(* IEC 61131-3 sources: PLC-IsaVODE/PLC-IsaVODE/samples/plc-programs, 701 files *)

(* ---- 250-building.IEC ---- *)
(*@PROPERTIES_EX@
TYPE: DATA_TYPE
LOCALE: 0
*)
(* ------------------------------------------- *)

TYPE oscat_TIMER_EVENT_DATA :
  STRUCT
	TYP          : BYTE;
	CHANNEL      : BYTE;
	DAY          : BYTE;
	START        : UDINT;
	DURATION     : TIME;
	LAND         : BYTE;
	LOR          : BYTE;
	LAST         : UDINT;
  END_STRUCT;
END_TYPE

TYPE
  oscat_TIMER_EVENT           : ARRAY [0..63]    OF oscat_TIMER_EVENT_DATA;
END_TYPE

(* ------------------------------------------- *)

TYPE
  oscat_T_AVG24         	  : ARRAY [0..47]   OF INT;

  oscat_TP4_qn                : ARRAY [0..3]    OF BOOL;

  oscat_bsa_X                 : ARRAY [0..2]    OF BYTE;
  oscat_blind_scene_array     : ARRAY [0..15]   OF oscat_bsa_X;

END_TYPE

(* ---- 731-WORLD_WEATHER.ST ---- *)
TYPE
  oscat_STRING30              : STRING;
  oscat_STRING250             : STRING;
  oscat_STRING8               : STRING;
  oscat_STRING60               : STRING;
  oscat_STRING3               : STRING;
  oscat_STRING10               : STRING;
END_TYPE

TYPE
  oscat_IP_FIFO128_DATA  : ARRAY [1..128] OF BYTE;
  oscat_Mailbox  : ARRAY [1..16] OF BYTE;

  oscat_IP_FIFO_DATA :
  STRUCT
	X       : oscat_IP_FIFO128_DATA; (* IP_ID FIFO Speicher          *)
	Y       : oscat_IP_FIFO128_DATA; (* IP_ID Z�hler                 *)
	ID      : BYTE;                  (* h�chste vergabene id         *)
	MAX_ID  : BYTE;                  (* maximal Anmeldungen pro ID   *)
    INIT    : BOOL;                  (* Initialisierung durchgef�hrt *)
	EMPTY   : BOOL;                  (* FIFO leer                    *)
	FULL    : BOOL;                  (* FIFO voll                    *)
	TOP     : INT;                   (* maximale anzahl in FIFO      *)
	NW      : INT;                   (* Schreibzeiger                *)
	NR      : INT;                   (* Lesezeiger                   *)
  END_STRUCT;

  oscat_IP_C:
  STRUCT
  	C_MODE:			BYTE;          		(*W Mode: TCP/UCP AKTIV/PASSIV                               *)
	C_PORT:         WORD;          		(*W Portnummer                                               *)
	C_IP:           DWORD;         		(*W IP-Adresse gepackt wwxxyyzz = www.xxx.yyy.zzz            *)
    C_STATE:        BYTE;          		(*R Verbindungsstatus ON/OFF + Flanke ON/OFF                 *)
	C_ENABLE:       BOOL;          		(*W Freigabe f�r Connect                                     *)
    R_OBSERVE:      BOOL;          		(*W Empfang ueberwachen                                      *)
    TIME_RESET:     BOOL;          		(*W Alle Timer ruecksetzen                                   *)
	ERROR:          DWORD;         		(*R vvwwxxyy (vv = CON_ERROR, ww = SEN_ERROR, xx = REC_ERROR *)
    FIFO:           oscat_IP_FIFO_DATA; (*I IP FIFO Struktur                                         *)
	MAILBOX:		oscat_Mailbox;		(*I Mailbox: Datenbereich f�r Bausteindatenaustausch         *)
  END_STRUCT;

  oscat_XML_CONTROL:
  STRUCT
    COMMAND:             WORD;            (*W                 *)
    WATCHDOG:            TIME;            (*W                 *)
    START_POS:           UINT;            (*W                 *)
    STOP_POS:            UINT;            (*W                 *)
    COUNT:               UINT;            (*R                 *)
    TYP:                 INT;             (*R                 *)
    LEVEL:               UINT;            (*R                 *)
    PATH:                oscat_STRING250; (*R                 *)
    ELEMENT:             oscat_STRING250; (*R                 *)
    ATTRIBUTE:           oscat_STRING250; (*R                 *)
    VALUE:               oscat_STRING250; (*R                 *)
    BLOCK1_START:        UINT;            (*R                 *)
    BLOCK1_STOP:         UINT;            (*R                 *)
    BLOCK2_START:        UINT;            (*R                 *)
    BLOCK2_STOP:         UINT;            (*R                 *)
  END_STRUCT;

  (* --------- WORLD WEATHER --------- *)

  oscat_WORLD_WEATHER_CUR :
  STRUCT
	OBSERVATION_TIME : oscat_STRING8;
	TEMP_C           : INT;
	WEATHER_CODE     : INT;
	WEATHER_DESC 	 : oscat_STRING60;
	WEATHER_ICON     : INT;
	WIND_SPEED_MILES : INT;
	WIND_SPEED_KMPH  : INT;
	WIND_DIR_DEGREE  : INT;
	WIND_DIR16POINT  : oscat_STRING3;
	PRECIPMM         : REAL;
	HUMIDITY         : INT;
	VISIBILITY       : INT;
	PRESSURE         : INT;
	CLOUDOVER        : INT;
  END_STRUCT;

  oscat_WORLD_WEATHER_DAY :
  STRUCT
	DATE_OF_DAY      : oscat_STRING10;
	TEMP_MAX_C       : INT;
	TEMP_MAX_F       : INT;
	TEMP_MIN_C       : INT;
	TEMP_MIN_F       : INT;
	WIND_SPEED_MILES : INT;
	WIND_SPEED_KMPH  : INT;
	WIND_DIR_DEGREE  : INT;
	WIND_DIR16POINT  : oscat_STRING3;
	WEATHER_CODE     : INT;
	WEATHER_DESC     : oscat_STRING60;
	WEATHER_ICON     : INT;
	PRECIPMM         : REAL;
  END_STRUCT;

  oscat_WORLD_WEATHER_DAY_ARR : ARRAY [0..4] OF oscat_WORLD_WEATHER_DAY;

  oscat_WORLD_WEATHER_DATA :
  STRUCT
	CUR : oscat_WORLD_WEATHER_CUR;
	DAY : oscat_WORLD_WEATHER_DAY_ARR;
  END_STRUCT;

  oscat_WORLD_WEATHER_aI0_41 : ARRAY[0..41] OF INT;

END_TYPE

TYPE
  oscat_NW_BUF_LONG  : ARRAY [0..4095] OF BYTE;

  oscat_NETWORK_BUFFER :
  STRUCT
    SIZE   : UINT;
    BUFFER : oscat_NW_BUF_LONG;
  END_STRUCT;

END_TYPE

FUNCTION_BLOCK WORLD_WEATHER_Block

	VAR_INPUT
		ACTIVATE :	BOOL;
		LATITUDE :	REAL;
		LONGITUDE :	REAL;
		KEY :	oscat_STRING30;
	END_VAR

	VAR_OUTPUT
		BUSY :	BOOL;
		DONE :	BOOL;
		ERROR_C :	DWORD;
		ERROR_T :	BYTE;
	END_VAR

	VAR_IN_OUT
		IP_C :	oscat_IP_C;
		S_BUF :	oscat_NETWORK_BUFFER;
		R_BUF :	oscat_NETWORK_BUFFER;
		WW :	oscat_WORLD_WEATHER_DATA;
	END_VAR

	VAR
		CHK_REAL :	CHK_REAL;
		REAL_TO_STRF :	REAL_TO_STRF;
		URL_DATA :	oscat_url;
		DNS_CLIENT :	DNS_CLIENT;
		HTTP_GET :	HTTP_GET;
		CPB :	CSV_PARSER_BUF;
		STRING_TO_URL :	STRING_TO_URL;
		FLOAT_TO_REAL :	FLOAT_TO_REAL;
		last_state :	BOOL;
		value_int :	INT;
		value_real :	REAL;
		v_real :	REAL;
		state :	INT;
		url_str :	oscat_STRING250;
		offset :	UDINT;
		size :	INT;
		sep :	BYTE;
		cnt :	INT;
		day :	INT;
		idx :	INT;
		run :	BYTE;
		result :	BYTE;
		value :	oscat_STRING250;
		DEC_TO_INT :	DEC_TO_INT;
		pos :	INT;
	END_VAR

	CASE state OF

	00:
		IF ACTIVATE AND NOT last_state THEN
			state := 20;
			DONE := FALSE;
			BUSY := TRUE;
			ERROR_C := DWORD#0;
			ERROR_T := BYTE#0;
		END_IF;

	20:
		REAL_TO_STRF(IN:=LATITUDE,N:=6,D:='.');
		url_str := CONCAT('http://free.worldweatheronline.com/feed/weather.ashx?q=',REAL_TO_STRF.REAL_TO_STRF);
		url_str := CONCAT(url_str,',');
		REAL_TO_STRF(IN:=LONGITUDE,N:=6,D:='.');
		url_str := CONCAT(url_str,REAL_TO_STRF.REAL_TO_STRF);
		url_str := CONCAT(url_str,'&format=csv&num_of_days=5&key=');
		url_str := CONCAT(url_str,key);

		STRING_TO_URL(STR:=url_str, DEFAULT_PROTOCOL:='', DEFAULT_PATH:='' );
		URL_DATA:=STRING_TO_URL.STRING_TO_URL;

		state := 40;

	40:
		IF DNS_CLIENT.DONE THEN
			state := 60;
		ELSIF (DNS_CLIENT.ERROR > DWORD#00) THEN
			ERROR_C := DNS_CLIENT.ERROR;
			ERROR_T := BYTE#01;
			state   := 100;
		END_IF;

	60:
		IF HTTP_GET.DONE THEN
			sep := BYTE#0;
			idx := 0;
			day := 0;
			cnt := 0;
			OFFSET := UINT_TO_UDINT(HTTP_GET.BODY_START);
			size := UINT_TO_INT(HTTP_GET.BODY_STOP);
			run := BYTE#1;
			state := 80;

		ELSIF (HTTP_GET.ERROR > DWORD#00) THEN
			ERROR_C := HTTP_GET.ERROR;
			ERROR_T := BYTE#02;
			state := 100;
		END_IF;

	80:	IF run = BYTE#0 THEN
			run := BYTE#1;
			IF result = BYTE#1 OR result = BYTE#2 THEN
				value_int := 0;
				value_real := 0.0;
				IF LEN(value) <= 20 THEN
					FLOAT_TO_REAL(FLT:=value);
					v_real := FLOAT_TO_REAL.FLOAT_TO_REAL;
					CHK_REAL(X := v_real);
					IF CHK_REAL.CHK_REAL = BYTE#0 THEN
						value_real := v_real;
						value_int := REAL_TO_INT(value_real);
					END_IF;
				END_IF;
				cnt := cnt + 1;
				IF cnt >=8 AND cnt <= 87 THEN
					IF cnt > 22 THEN
						CASE idx OF
						00:	WW.DAY[day].DATE_OF_DAY := value;
						01:	WW.DAY[day].TEMP_MAX_C := value_int;
						02:	WW.DAY[day].TEMP_MAX_F := value_int;
						03:	WW.DAY[day].TEMP_MIN_C := value_int;
						04:	WW.DAY[day].TEMP_MIN_F := value_int;
						05:	WW.DAY[day].WIND_SPEED_MILES := value_int;
						06:	WW.DAY[day].WIND_SPEED_KMPH := value_int;
						07:	WW.DAY[day].WIND_DIR_DEGREE := value_int;
						08:	WW.DAY[day].WIND_DIR16POINT := value;
						09:	WW.DAY[day].WEATHER_CODE := value_int;
						10:	pos := FIND(value, '/wsymbol_');
							IF pos > 0 AND LEN(value) > pos + 13 THEN
								DEC_TO_INT(DEC:=MID(value,4,pos + 9));
								WW.DAY[day].WEATHER_ICON := DEC_TO_INT.DEC_TO_INT;
							ELSE
								WW.DAY[day].WEATHER_ICON := 0;
							END_IF;
						11:	WW.DAY[day].WEATHER_DESC := value;
						12:	WW.DAY[day].PRECIPMM := value_real;
						END_CASE;
						idx := idx + 1;
						IF idx > 12 THEN
							idx := 0;
							day := day + 1;
						END_IF;
					ELSE
						CASE cnt OF
						08:	sep := BYTE#44;
						09:	WW.CUR.OBSERVATION_TIME := value;
						10:	WW.CUR.TEMP_C := value_int;
						11:	WW.CUR.WEATHER_CODE := value_int;
						12:	pos := FIND(value, '/wsymbol_');
							IF pos > 0 AND LEN(value) > pos + 13 THEN
								DEC_TO_INT(DEC:=MID(value,4,pos + 9));
								WW.CUR.WEATHER_ICON := DEC_TO_INT.DEC_TO_INT;
							ELSE
								WW.CUR.WEATHER_ICON := 0;
							END_IF;
						13:	WW.CUR.WEATHER_DESC := value;
						14:	WW.CUR.WIND_SPEED_MILES := value_int;
						15:	WW.CUR.WIND_SPEED_KMPH := value_int;
						16:	WW.CUR.WIND_DIR_DEGREE := value_int;
						17:	WW.CUR.WIND_DIR16POINT := value;
						18:	WW.CUR.PRECIPMM := value_real;
						19:	WW.CUR.HUMIDITY := value_int;
						20:	WW.CUR.VISIBILITY := value_int;
						21:	WW.CUR.PRESSURE := value_int;
						22:	WW.CUR.CLOUDOVER := value_int;
						END_CASE;
					END_IF;
				END_IF;
			ELSIF result = BYTE#10 THEN
				DONE  := TRUE;
				run := BYTE#0;
				state := 100;
			END_IF;
		END_IF;

	100:
		IF (NOT HTTP_GET.DONE) THEN
			state := 0;
			BUSY := FALSE;
			DONE := ERROR_T = BYTE#0;
		END_IF;

	END_CASE;

	DNS_CLIENT.IP_C     := IP_C;
	DNS_CLIENT.S_BUF    := S_BUF;
	DNS_CLIENT.R_BUF    := R_BUF;
	DNS_CLIENT.DOMAIN   := URL_DATA.DOMAIN;
	DNS_CLIENT.IP4_DNS  := DWORD#00;
	DNS_CLIENT.ACTIVATE := state=40;
	DNS_CLIENT();
	IP_C  := DNS_CLIENT.IP_C;
	S_BUF := DNS_CLIENT.S_BUF;
	R_BUF := DNS_CLIENT.R_BUF;

	HTTP_GET.IP_C        := IP_C;
	HTTP_GET.S_BUF       := S_BUF;
	HTTP_GET.R_BUF       := R_BUF;
	HTTP_GET.IP4         := DNS_CLIENT.IP4;
	HTTP_GET.GET         := state=60;
	HTTP_GET.MODE        := BYTE#2;
	HTTP_GET.UNLOCK_BUF  := state=100;
	HTTP_GET.URL_DATA    := URL_DATA;
	HTTP_GET();
	IP_C     := HTTP_GET.IP_C;
	S_BUF    := HTTP_GET.S_BUF;
	R_BUF    := HTTP_GET.R_BUF;
	URL_DATA := HTTP_GET.URL_DATA;

	CPB(SEP:=sep,RUN:=run,OFFSET:=offset,VALUE:=value,PT:=R_BUF);
	run:=CPB.RUN;
	offset:=CPB.OFFSET;
	value:=CPB.VALUE;
	R_BUF:=CPB.PT;
	result:=CPB.RESULT;

	last_state := ACTIVATE;

END_FUNCTION_BLOCK

PROGRAM program0
	VAR
		ACTIVATE :	BOOL;
		LATITUDE :	REAL;
		LONGITUDE :	REAL;
		KEY :	oscat_STRING30;
		IP_C :	oscat_IP_C;
		S_BUF :	oscat_NETWORK_BUFFER;
		R_BUF :	oscat_NETWORK_BUFFER;
		WW :	oscat_WORLD_WEATHER_DATA;
		BUSY :	BOOL;
		DONE :	BOOL;
		ERROR_C :	DWORD;
		ERROR_T :	BYTE;

		func_block : WORLD_WEATHER_Block;
	END_VAR
	func_block.ACTIVATE := ACTIVATE;
	func_block.LATITUDE := LATITUDE;
	func_block.LONGITUDE := LONGITUDE;
	func_block.KEY := KEY;
	func_block.IP_C := IP_C;
	func_block.S_BUF := S_BUF;
	func_block.R_BUF := R_BUF;
	func_block.WW := WW;

	func_block();
	IP_C  := func_block.IP_C;
	S_BUF  := func_block.S_BUF;
	R_BUF  := func_block.R_BUF;
	WW  := func_block.WW;
	BUSY  := func_block.BUSY;
	DONE  := func_block.DONE;
	ERROR_C  := func_block.ERROR_C;
	ERROR_T  := func_block.ERROR_T;
END_PROGRAM

CONFIGURATION Config0
	RESOURCE Res0 ON PLC
		TASK task0(INTERVAL := T#20ms,PRIORITY := 0);
		PROGRAM instance0 WITH task0 : program0;
	END_RESOURCE
END_CONFIGURATION

(* ---- 733-YAHOO_WEATHER_ICON_OSCAT.ST ---- *)
TYPE
  oscat_STRING1               : STRING;
  oscat_STRING2               : STRING;
  oscat_STRING3               : STRING;
  oscat_STRING4               : STRING;
  oscat_STRING5               : STRING;
  oscat_STRING8               : STRING;
  oscat_STRING10              : STRING;
  oscat_STRING12            : STRING;
  oscat_STRING15            : STRING;
  oscat_STRING20            : STRING;
  oscat_STRING27            : STRING;
  oscat_STRING30            : STRING;
  oscat_STRING32            : STRING;
  oscat_STRING40            : STRING;
  oscat_STRING48            : STRING;
  oscat_STRING50            : STRING;
  oscat_STRING60            : STRING;
  oscat_STRING64            : STRING;
  oscat_STRING80            : STRING;
  oscat_STRING120            : STRING;
  oscat_STRING140            : STRING;
  oscat_STRING160            : STRING;
  oscat_STRING180            : STRING;
  oscat_STRING190            : STRING;
  oscat_STRING250            : STRING;
END_TYPE

TYPE
  oscat_IP_FIFO128_DATA  : ARRAY [1..128] OF BYTE;
  oscat_Mailbox  : ARRAY [1..16] OF BYTE;

  oscat_IP_FIFO_DATA :
  STRUCT
	X       : oscat_IP_FIFO128_DATA; (* IP_ID FIFO Speicher          *)
	Y       : oscat_IP_FIFO128_DATA; (* IP_ID Z�hler                 *)
	ID      : BYTE;                  (* h�chste vergabene id         *)
	MAX_ID  : BYTE;                  (* maximal Anmeldungen pro ID   *)
    INIT    : BOOL;                  (* Initialisierung durchgef�hrt *)
	EMPTY   : BOOL;                  (* FIFO leer                    *)
	FULL    : BOOL;                  (* FIFO voll                    *)
	TOP     : INT;                   (* maximale anzahl in FIFO      *)
	NW      : INT;                   (* Schreibzeiger                *)
	NR      : INT;                   (* Lesezeiger                   *)
  END_STRUCT;

  oscat_IP_C:
  STRUCT
  	C_MODE:			BYTE;          		(*W Mode: TCP/UCP AKTIV/PASSIV                               *)
	C_PORT:         WORD;          		(*W Portnummer                                               *)
	C_IP:           DWORD;         		(*W IP-Adresse gepackt wwxxyyzz = www.xxx.yyy.zzz            *)
    C_STATE:        BYTE;          		(*R Verbindungsstatus ON/OFF + Flanke ON/OFF                 *)
	C_ENABLE:       BOOL;          		(*W Freigabe f�r Connect                                     *)
    R_OBSERVE:      BOOL;          		(*W Empfang ueberwachen                                      *)
    TIME_RESET:     BOOL;          		(*W Alle Timer ruecksetzen                                   *)
	ERROR:          DWORD;         		(*R vvwwxxyy (vv = CON_ERROR, ww = SEN_ERROR, xx = REC_ERROR *)
    FIFO:           oscat_IP_FIFO_DATA; (*I IP FIFO Struktur                                         *)
	MAILBOX:		oscat_Mailbox;		(*I Mailbox: Datenbereich f�r Bausteindatenaustausch         *)
  END_STRUCT;

  oscat_XML_CONTROL:
  STRUCT
    COMMAND:             WORD;            (*W                 *)
    WATCHDOG:            TIME;            (*W                 *)
    START_POS:           UINT;            (*W                 *)
    STOP_POS:            UINT;            (*W                 *)
    COUNT:               UINT;            (*R                 *)
    TYP:                 INT;             (*R                 *)
    LEVEL:               UINT;            (*R                 *)
    PATH:                oscat_STRING250; (*R                 *)
    ELEMENT:             oscat_STRING250; (*R                 *)
    ATTRIBUTE:           oscat_STRING250; (*R                 *)
    VALUE:               oscat_STRING250; (*R                 *)
    BLOCK1_START:        UINT;            (*R                 *)
    BLOCK1_STOP:         UINT;            (*R                 *)
    BLOCK2_START:        UINT;            (*R                 *)
    BLOCK2_STOP:         UINT;            (*R                 *)
  END_STRUCT;

  (* --------- WORLD WEATHER --------- *)

  oscat_WORLD_WEATHER_CUR :
  STRUCT
	OBSERVATION_TIME : oscat_STRING8;
	TEMP_C           : INT;
	WEATHER_CODE     : INT;
	WEATHER_DESC 	 : oscat_STRING60;
	WEATHER_ICON     : INT;
	WIND_SPEED_MILES : INT;
	WIND_SPEED_KMPH  : INT;
	WIND_DIR_DEGREE  : INT;
	WIND_DIR16POINT  : oscat_STRING3;
	PRECIPMM         : REAL;
	HUMIDITY         : INT;
	VISIBILITY       : INT;
	PRESSURE         : INT;
	CLOUDOVER        : INT;
  END_STRUCT;

  oscat_WORLD_WEATHER_DAY :
  STRUCT
	DATE_OF_DAY      : oscat_STRING10;
	TEMP_MAX_C       : INT;
	TEMP_MAX_F       : INT;
	TEMP_MIN_C       : INT;
	TEMP_MIN_F       : INT;
	WIND_SPEED_MILES : INT;
	WIND_SPEED_KMPH  : INT;
	WIND_DIR_DEGREE  : INT;
	WIND_DIR16POINT  : oscat_STRING3;
	WEATHER_CODE     : INT;
	WEATHER_DESC     : oscat_STRING60;
	WEATHER_ICON     : INT;
	PRECIPMM         : REAL;
  END_STRUCT;

  oscat_WORLD_WEATHER_DAY_ARR : ARRAY [0..4] OF oscat_WORLD_WEATHER_DAY;

  oscat_WORLD_WEATHER_DATA :
  STRUCT
	CUR : oscat_WORLD_WEATHER_CUR;
	DAY : oscat_WORLD_WEATHER_DAY_ARR;
  END_STRUCT;

  oscat_WORLD_WEATHER_aI0_41 : ARRAY[0..41] OF INT;

  (* --------- WEATHER CHANNEL --------- *)
  oscat_YAHOO_WEATHER_DATA:
  STRUCT
    TIMETOLIVE:                 INT;              (* TIME TO LIVE: HOW LONG IN MINUTES THIS FEED SHOULD BE CACHED         *)
    LOCATION_CITY:              OSCAT_STRING40;   (* THE LOCATION OF THIS FORECAST: CITY: CITY NAME  *)
    LOCATION_REGION:            OSCAT_STRING20;   (* THE LOCATION OF THIS FORECAST: REGION: STATE, TERRITORY, OR REGION, IF GIVEN *)
    LOCATION_COUNTRY:           OSCAT_STRING20;    (* THE LOCATION OF THIS FORECAST: COUNTRY: TWO-CHARACTER COUNTRY CODE *)
    UNIT_TEMPERATURE:           OSCAT_STRING1;    (* TEMPERATURE: DEGREE UNITS, F FOR FAHRENHEIT OR C FOR CELSIUS *)
    UNIT_DISTANCE:              OSCAT_STRING2;    (* DISTANCE: UNITS FOR DISTANCE, MI FOR MILES OR KM FOR KILOMETERS *)
    UNIT_PRESSURE:              OSCAT_STRING2;    (* PRESSURE: UNITS OF BAROMETRIC PRESSURE, IN FOR POUNDS PER SQUARE INCH OR MB FOR MILLIBARS *)
    UNIT_SPEED:                 OSCAT_STRING4;    (* SPEED: UNITS OF SPEED, MPH FOR MILES PER HOUR OR KPH FOR KILOMETERS PER HOUR *)
    WIND_CHILL:                 INT;              (* FORECAST INFORMATION ABOUT WIND CHILL IN DEGREES *)
    WIND_DIRECTION:             INT;              (* FORECAST INFORMATION ABOUT WIND DIRECTION, IN DEGREES *)
    WIND_SPEED:                 REAL;             (* FORECAST INFORMATION ABOUT WIND SPEED, IN THE UNITS (MPH OR KPH)*)
    ATMOSPHERE_HUMIDITY:        INT;              (* FORECAST INFORMATION ABOUT CURRENT ATMOSPHERIC HUMIDITY: HUMIDITY, IN PERCENT  *)
    ATMOSPHERE_PRESSURE:        INT;              (* FORECAST INFORMATION ABOUT CURRENT ATMOSPHERIC PRESSURE: BAROMETRIC PRESSURE, IN THE UNITS (IN OR MB) *)
	ATMOSPHERE_VISIBILITY:      REAL;             (* FORECAST INFORMATION ABOUT CURRENT ATMOSPHERIC VISIBILITY, IN THE UNITS (MI OR KM) *)
	ATMOSPHERE_RISING:          INT;              (* FORECAST INFORMATION ABOUT RISING: STATE OF THE BAROMETRIC PRESSURE: STEADY (0), RISING (1), OR FALLING (2). (INTEGER: 0, 1, 2) *)
    ASTRONOMY_SUNRISE:          OSCAT_STRING10;   (* SUNRISE: TODAY'S SUNRISE TIME. THE TIME IS A STRING IN A LOCAL TIME FORMAT OF "H:MM AM/PM" *)
    ASTRONOMY_SUNSET:           OSCAT_STRING10;   (* SUNSET: TODAY'S SUNSET TIME. THE TIME IS A STRING IN A LOCAL TIME FORMAT OF "H:MM AM/PM", *)
    GEO_LATITUDE:               REAL;             (* THE LATITUDE OF THE LOCATION *)
    GEO_LONGITUDE:              REAL;             (* THE LONGITUDE OF THE LOCATION *)
    CUR_CONDITIONS_TEMP:        INT;              (* THE CURRENT WEATHER CONDITIONS: TEMP: THE CURRENT TEMPERATURE, IN THE UNITS (F OR C) *)
    CUR_CONDITIONS_TEXT:        OSCAT_STRING40;   (* THE CURRENT WEATHER CONDITIONS: TEXT: A TEXTUAL DESCRIPTION OF CONDITIONS *)
    CUR_CONDITIONS_CODE:        INT;              (* THE CURRENT WEATHER CONDITIONS: CODE: THE CONDITION CODE FOR THIS FORECAST *)
	CUR_CONDITIONS_ICON:        INT;			  (* THE CURRENT WEATHER CONDITIONS: ICON: THE CONDITION ICON FOR THIS FORECAST *)
    FORCAST_TODAY_LOW_TEMP:     INT;              (* THE FORCAST TODAY WEATHER CONDITIONS: THE FORECASTED LOW TEMPERATURE FOR THIS DAY IN THE UNITS (F OR C) *)
    FORCAST_TODAY_HIGH_TEMP:    INT;              (* THE FORCAST TODAY WEATHER CONDITIONS: THE FORECASTED HIGH TEMPERATURE FOR THIS DAY IN THE UNITS (F OR C) *)
    FORCAST_TODAY_TEXT:         OSCAT_STRING40;   (* THE FORCAST TODAY WEATHER CONDITIONS: TEXT: A TEXTUAL DESCRIPTION OF CONDITIONS *)
    FORCAST_TODAY_CODE:         INT;              (* THE CURRENT WEATHER CONDITIONS: CODE: THE CONDITION CODE FOR THIS FORECAST *)
	FORCAST_TODAY_ICON:         INT;			  (* THE CURRENT WEATHER CONDITIONS: ICON: THE CONDITION ICON FOR THIS FORECAST *)
    FORCAST_TOMORROW_LOW_TEMP:  INT;              (* THE FORCAST TOMORROW WEATHER CONDITIONS: THE FORECASTED LOW TEMPERATURE FOR THIS DAY IN THE UNITS (F OR C) *)
    FORCAST_TOMORROW_HIGH_TEMP: INT;              (* THE FORCAST TOMORROW WEATHER CONDITIONS: THE FORECASTED HIGH TEMPERATURE FOR THIS DAY IN THE UNITS (F OR C) *)
    FORCAST_TOMORROW_TEXT:      OSCAT_STRING40;   (* THE FORCAST TOMORROW WEATHER CONDITIONS: TEXT: A TEXTUAL DESCRIPTION OF CONDITIONS *)
    FORCAST_TOMORROW_CODE:      INT;              (* THE CURRENT WEATHER CONDITIONS: CODE: THE CONDITION CODE FOR THIS FORECAST *)
	FORCAST_TOMORROW_ICON:      INT;			  (* THE CURRENT WEATHER CONDITIONS: ICON: THE CONDITION ICON FOR THIS FORECAST *)
  END_STRUCT;

  oscat_YAHOO_WEATHER_aI0_48 : ARRAY[0..48] OF INT;

  oscat_IP2GEO_DATA:
  STRUCT
	STATE :				BOOL;			  (* STATE *)
	IP4 :				DWORD;			  (* IP-Adresse *)
    COUNTRY_CODE :		oscat_STRING2;    (*   *)
    COUNTRY_NAME :		oscat_STRING20;   (*   *)
    REGION_CODE :		oscat_STRING2;    (*   *)
    REGION_NAME :		oscat_STRING20;   (*   *)
    CITY :				oscat_STRING20;   (*   *)
    GEO_LATITUDE :		REAL;             (*   *)
    GEO_LONGITUDE :		REAL;             (*   *)
	TIME_ZONE_NAME :	oscat_STRING20;
	GMT_OFFSET :		INT;
	IS_DST :			BOOL;
  END_STRUCT;
END_TYPE

FUNCTION_BLOCK YAHOO_WEATHER_ICON_OSCAT_Block

	VAR_INPUT
		ACTIVATE :	BOOL;
	END_VAR

	VAR_IN_OUT
		YW :	oscat_YAHOO_WEATHER_DATA;
	END_VAR

	VAR
		act_last :	BOOL;
		x :	INT;
		init :	BOOL;
		dat :	oscat_YAHOO_WEATHER_aI0_48;
	END_VAR

	IF not init THEN
		init := TRUE;

		dat[00] := 4;
		dat[01] := 2;
		dat[02] := 2;
		dat[03] := 4;
		dat[04] := 17;
		dat[05] := 1;
		dat[06] := 3;
		dat[07] := 1;
		dat[08] := 2;
		dat[09] := 2;
		dat[10] := 2;
		dat[11] := 2;
		dat[12] := 2;
		dat[13] := 3;
		dat[14] := 3;
		dat[15] := 3;
		dat[16] := 3;
		dat[17] := 5;
		dat[18] := 3;
		dat[19] := 6;
		dat[20] := 7;
		dat[21] := 14;
		dat[22] := 8;
		dat[23] := 9;
		dat[24] := 9;
		dat[25] := 10;
		dat[26] := 9;
		dat[27] := 11;
		dat[28] := 12;
		dat[29] := 11;
		dat[30] := 12;
		dat[31] := 13;
		dat[32] := 14;
		dat[33] := 15;
		dat[34] := 16;
		dat[35] := 4;
		dat[36] := 14;
		dat[37] := 4;
		dat[38] := 17;
		dat[39] := 2;
		dat[40] := 2;
		dat[41] := 3;
		dat[42] := 3;
		dat[43] := 3;
		dat[44] := 12;
		dat[45] := 2;
		dat[46] := 3;
		dat[47] := 4;
		dat[48] := 0;
	END_IF;

	IF ACTIVATE AND act_last = FALSE THEN
		x := MIN(YW.CUR_CONDITIONS_CODE,48);
		YW.CUR_CONDITIONS_ICON := dat[x];
		x := MIN(YW.FORCAST_TODAY_CODE,48);
		YW.FORCAST_TODAY_ICON := dat[x];
		x := MIN(YW.FORCAST_TOMORROW_CODE,48);
		YW.FORCAST_TOMORROW_ICON := dat[x];
	END_IF;
	act_last := ACTIVATE;

END_FUNCTION_BLOCK

PROGRAM program0
	VAR
		ACTIVATE :	BOOL;
		YW :	oscat_YAHOO_WEATHER_DATA;

		func_block : YAHOO_WEATHER_ICON_OSCAT_Block;
	END_VAR
	func_block.ACTIVATE := ACTIVATE;
	func_block.YW := YW;

	func_block();
	YW  := func_block.YW;
END_PROGRAM

CONFIGURATION Config0
	RESOURCE Res0 ON PLC
		TASK task0(INTERVAL := T#20ms,PRIORITY := 0);
		PROGRAM instance0 WITH task0 : program0;
	END_RESOURCE
END_CONFIGURATION

(* ---- 737-YAHOO_WEATHER_DESC_GE.ST ---- *)
TYPE
  oscat_STRING1               : STRING;
  oscat_STRING2               : STRING;
  oscat_STRING3               : STRING;
  oscat_STRING4               : STRING;
  oscat_STRING5               : STRING;
  oscat_STRING8               : STRING;
  oscat_STRING10              : STRING;
  oscat_STRING12            : STRING;
  oscat_STRING15            : STRING;
  oscat_STRING20            : STRING;
  oscat_STRING27            : STRING;
  oscat_STRING30            : STRING;
  oscat_STRING32            : STRING;
  oscat_STRING40            : STRING;
  oscat_STRING48            : STRING;
  oscat_STRING50            : STRING;
  oscat_STRING60            : STRING;
  oscat_STRING64            : STRING;
  oscat_STRING80            : STRING;
  oscat_STRING120            : STRING;
  oscat_STRING140            : STRING;
  oscat_STRING160            : STRING;
  oscat_STRING180            : STRING;
  oscat_STRING190            : STRING;
  oscat_STRING250            : STRING;
END_TYPE

TYPE
  oscat_IP_FIFO128_DATA  : ARRAY [1..128] OF BYTE;
  oscat_Mailbox  : ARRAY [1..16] OF BYTE;

  oscat_IP_FIFO_DATA :
  STRUCT
	X       : oscat_IP_FIFO128_DATA; (* IP_ID FIFO Speicher          *)
	Y       : oscat_IP_FIFO128_DATA; (* IP_ID Z�hler                 *)
	ID      : BYTE;                  (* h�chste vergabene id         *)
	MAX_ID  : BYTE;                  (* maximal Anmeldungen pro ID   *)
    INIT    : BOOL;                  (* Initialisierung durchgef�hrt *)
	EMPTY   : BOOL;                  (* FIFO leer                    *)
	FULL    : BOOL;                  (* FIFO voll                    *)
	TOP     : INT;                   (* maximale anzahl in FIFO      *)
	NW      : INT;                   (* Schreibzeiger                *)
	NR      : INT;                   (* Lesezeiger                   *)
  END_STRUCT;

  oscat_IP_C:
  STRUCT
  	C_MODE:			BYTE;          		(*W Mode: TCP/UCP AKTIV/PASSIV                               *)
	C_PORT:         WORD;          		(*W Portnummer                                               *)
	C_IP:           DWORD;         		(*W IP-Adresse gepackt wwxxyyzz = www.xxx.yyy.zzz            *)
    C_STATE:        BYTE;          		(*R Verbindungsstatus ON/OFF + Flanke ON/OFF                 *)
	C_ENABLE:       BOOL;          		(*W Freigabe f�r Connect                                     *)
    R_OBSERVE:      BOOL;          		(*W Empfang ueberwachen                                      *)
    TIME_RESET:     BOOL;          		(*W Alle Timer ruecksetzen                                   *)
	ERROR:          DWORD;         		(*R vvwwxxyy (vv = CON_ERROR, ww = SEN_ERROR, xx = REC_ERROR *)
    FIFO:           oscat_IP_FIFO_DATA; (*I IP FIFO Struktur                                         *)
	MAILBOX:		oscat_Mailbox;		(*I Mailbox: Datenbereich f�r Bausteindatenaustausch         *)
  END_STRUCT;

  oscat_XML_CONTROL:
  STRUCT
    COMMAND:             WORD;            (*W                 *)
    WATCHDOG:            TIME;            (*W                 *)
    START_POS:           UINT;            (*W                 *)
    STOP_POS:            UINT;            (*W                 *)
    COUNT:               UINT;            (*R                 *)
    TYP:                 INT;             (*R                 *)
    LEVEL:               UINT;            (*R                 *)
    PATH:                oscat_STRING250; (*R                 *)
    ELEMENT:             oscat_STRING250; (*R                 *)
    ATTRIBUTE:           oscat_STRING250; (*R                 *)
    VALUE:               oscat_STRING250; (*R                 *)
    BLOCK1_START:        UINT;            (*R                 *)
    BLOCK1_STOP:         UINT;            (*R                 *)
    BLOCK2_START:        UINT;            (*R                 *)
    BLOCK2_STOP:         UINT;            (*R                 *)
  END_STRUCT;

  (* --------- WORLD WEATHER --------- *)

  oscat_WORLD_WEATHER_CUR :
  STRUCT
	OBSERVATION_TIME : oscat_STRING8;
	TEMP_C           : INT;
	WEATHER_CODE     : INT;
	WEATHER_DESC 	 : oscat_STRING60;
	WEATHER_ICON     : INT;
	WIND_SPEED_MILES : INT;
	WIND_SPEED_KMPH  : INT;
	WIND_DIR_DEGREE  : INT;
	WIND_DIR16POINT  : oscat_STRING3;
	PRECIPMM         : REAL;
	HUMIDITY         : INT;
	VISIBILITY       : INT;
	PRESSURE         : INT;
	CLOUDOVER        : INT;
  END_STRUCT;

  oscat_WORLD_WEATHER_DAY :
  STRUCT
	DATE_OF_DAY      : oscat_STRING10;
	TEMP_MAX_C       : INT;
	TEMP_MAX_F       : INT;
	TEMP_MIN_C       : INT;
	TEMP_MIN_F       : INT;
	WIND_SPEED_MILES : INT;
	WIND_SPEED_KMPH  : INT;
	WIND_DIR_DEGREE  : INT;
	WIND_DIR16POINT  : oscat_STRING3;
	WEATHER_CODE     : INT;
	WEATHER_DESC     : oscat_STRING60;
	WEATHER_ICON     : INT;
	PRECIPMM         : REAL;
  END_STRUCT;

  oscat_WORLD_WEATHER_DAY_ARR : ARRAY [0..4] OF oscat_WORLD_WEATHER_DAY;

  oscat_WORLD_WEATHER_DATA :
  STRUCT
	CUR : oscat_WORLD_WEATHER_CUR;
	DAY : oscat_WORLD_WEATHER_DAY_ARR;
  END_STRUCT;

  oscat_WORLD_WEATHER_aI0_41 : ARRAY[0..41] OF INT;

  (* --------- WEATHER CHANNEL --------- *)
  oscat_YAHOO_WEATHER_DATA:
  STRUCT
    TIMETOLIVE:                 INT;              (* TIME TO LIVE: HOW LONG IN MINUTES THIS FEED SHOULD BE CACHED         *)
    LOCATION_CITY:              OSCAT_STRING40;   (* THE LOCATION OF THIS FORECAST: CITY: CITY NAME  *)
    LOCATION_REGION:            OSCAT_STRING20;   (* THE LOCATION OF THIS FORECAST: REGION: STATE, TERRITORY, OR REGION, IF GIVEN *)
    LOCATION_COUNTRY:           OSCAT_STRING20;    (* THE LOCATION OF THIS FORECAST: COUNTRY: TWO-CHARACTER COUNTRY CODE *)
    UNIT_TEMPERATURE:           OSCAT_STRING1;    (* TEMPERATURE: DEGREE UNITS, F FOR FAHRENHEIT OR C FOR CELSIUS *)
    UNIT_DISTANCE:              OSCAT_STRING2;    (* DISTANCE: UNITS FOR DISTANCE, MI FOR MILES OR KM FOR KILOMETERS *)
    UNIT_PRESSURE:              OSCAT_STRING2;    (* PRESSURE: UNITS OF BAROMETRIC PRESSURE, IN FOR POUNDS PER SQUARE INCH OR MB FOR MILLIBARS *)
    UNIT_SPEED:                 OSCAT_STRING4;    (* SPEED: UNITS OF SPEED, MPH FOR MILES PER HOUR OR KPH FOR KILOMETERS PER HOUR *)
    WIND_CHILL:                 INT;              (* FORECAST INFORMATION ABOUT WIND CHILL IN DEGREES *)
    WIND_DIRECTION:             INT;              (* FORECAST INFORMATION ABOUT WIND DIRECTION, IN DEGREES *)
    WIND_SPEED:                 REAL;             (* FORECAST INFORMATION ABOUT WIND SPEED, IN THE UNITS (MPH OR KPH)*)
    ATMOSPHERE_HUMIDITY:        INT;              (* FORECAST INFORMATION ABOUT CURRENT ATMOSPHERIC HUMIDITY: HUMIDITY, IN PERCENT  *)
    ATMOSPHERE_PRESSURE:        INT;              (* FORECAST INFORMATION ABOUT CURRENT ATMOSPHERIC PRESSURE: BAROMETRIC PRESSURE, IN THE UNITS (IN OR MB) *)
	ATMOSPHERE_VISIBILITY:      REAL;             (* FORECAST INFORMATION ABOUT CURRENT ATMOSPHERIC VISIBILITY, IN THE UNITS (MI OR KM) *)
	ATMOSPHERE_RISING:          INT;              (* FORECAST INFORMATION ABOUT RISING: STATE OF THE BAROMETRIC PRESSURE: STEADY (0), RISING (1), OR FALLING (2). (INTEGER: 0, 1, 2) *)
    ASTRONOMY_SUNRISE:          OSCAT_STRING10;   (* SUNRISE: TODAY'S SUNRISE TIME. THE TIME IS A STRING IN A LOCAL TIME FORMAT OF "H:MM AM/PM" *)
    ASTRONOMY_SUNSET:           OSCAT_STRING10;   (* SUNSET: TODAY'S SUNSET TIME. THE TIME IS A STRING IN A LOCAL TIME FORMAT OF "H:MM AM/PM", *)
    GEO_LATITUDE:               REAL;             (* THE LATITUDE OF THE LOCATION *)
    GEO_LONGITUDE:              REAL;             (* THE LONGITUDE OF THE LOCATION *)
    CUR_CONDITIONS_TEMP:        INT;              (* THE CURRENT WEATHER CONDITIONS: TEMP: THE CURRENT TEMPERATURE, IN THE UNITS (F OR C) *)
    CUR_CONDITIONS_TEXT:        OSCAT_STRING40;   (* THE CURRENT WEATHER CONDITIONS: TEXT: A TEXTUAL DESCRIPTION OF CONDITIONS *)
    CUR_CONDITIONS_CODE:        INT;              (* THE CURRENT WEATHER CONDITIONS: CODE: THE CONDITION CODE FOR THIS FORECAST *)
	CUR_CONDITIONS_ICON:        INT;			  (* THE CURRENT WEATHER CONDITIONS: ICON: THE CONDITION ICON FOR THIS FORECAST *)
    FORCAST_TODAY_LOW_TEMP:     INT;              (* THE FORCAST TODAY WEATHER CONDITIONS: THE FORECASTED LOW TEMPERATURE FOR THIS DAY IN THE UNITS (F OR C) *)
    FORCAST_TODAY_HIGH_TEMP:    INT;              (* THE FORCAST TODAY WEATHER CONDITIONS: THE FORECASTED HIGH TEMPERATURE FOR THIS DAY IN THE UNITS (F OR C) *)
    FORCAST_TODAY_TEXT:         OSCAT_STRING40;   (* THE FORCAST TODAY WEATHER CONDITIONS: TEXT: A TEXTUAL DESCRIPTION OF CONDITIONS *)
    FORCAST_TODAY_CODE:         INT;              (* THE CURRENT WEATHER CONDITIONS: CODE: THE CONDITION CODE FOR THIS FORECAST *)
	FORCAST_TODAY_ICON:         INT;			  (* THE CURRENT WEATHER CONDITIONS: ICON: THE CONDITION ICON FOR THIS FORECAST *)
    FORCAST_TOMORROW_LOW_TEMP:  INT;              (* THE FORCAST TOMORROW WEATHER CONDITIONS: THE FORECASTED LOW TEMPERATURE FOR THIS DAY IN THE UNITS (F OR C) *)
    FORCAST_TOMORROW_HIGH_TEMP: INT;              (* THE FORCAST TOMORROW WEATHER CONDITIONS: THE FORECASTED HIGH TEMPERATURE FOR THIS DAY IN THE UNITS (F OR C) *)
    FORCAST_TOMORROW_TEXT:      OSCAT_STRING40;   (* THE FORCAST TOMORROW WEATHER CONDITIONS: TEXT: A TEXTUAL DESCRIPTION OF CONDITIONS *)
    FORCAST_TOMORROW_CODE:      INT;              (* THE CURRENT WEATHER CONDITIONS: CODE: THE CONDITION CODE FOR THIS FORECAST *)
	FORCAST_TOMORROW_ICON:      INT;			  (* THE CURRENT WEATHER CONDITIONS: ICON: THE CONDITION ICON FOR THIS FORECAST *)
  END_STRUCT;

  oscat_YAHOO_WEATHER_aI0_48 : ARRAY[0..48] OF INT;

  oscat_IP2GEO_DATA:
  STRUCT
	STATE :				BOOL;			  (* STATE *)
	IP4 :				DWORD;			  (* IP-Adresse *)
    COUNTRY_CODE :		oscat_STRING2;    (*   *)
    COUNTRY_NAME :		oscat_STRING20;   (*   *)
    REGION_CODE :		oscat_STRING2;    (*   *)
    REGION_NAME :		oscat_STRING20;   (*   *)
    CITY :				oscat_STRING20;   (*   *)
    GEO_LATITUDE :		REAL;             (*   *)
    GEO_LONGITUDE :		REAL;             (*   *)
	TIME_ZONE_NAME :	oscat_STRING20;
	GMT_OFFSET :		INT;
	IS_DST :			BOOL;
  END_STRUCT;
END_TYPE

FUNCTION_BLOCK YAHOO_WEATHER_DESC_GE_Block

	VAR_INPUT
		ACTIVATE :	BOOL;
	END_VAR

	VAR_IN_OUT
		YW :	oscat_YAHOO_WEATHER_DATA;
	END_VAR

	VAR
		act_last :	BOOL;
		x :	INT;
		y :	INT;
		str :	oscat_STRING40;
	END_VAR

	IF ACTIVATE AND act_last = FALSE THEN
		FOR y := 1 TO 4 DO
			CASE y OF
			1:	x := YW.CUR_CONDITIONS_CODE;
			2 :	YW.CUR_CONDITIONS_TEXT := str;
				x := YW.FORCAST_TODAY_CODE;
			3 :	YW.FORCAST_TODAY_TEXT := str;
				x := YW.FORCAST_TOMORROW_CODE;
			4 :	YW.FORCAST_TOMORROW_TEXT := str;
			END_CASE;

			CASE x OF
			00:	str := 'Wirbelsturm';
			01:	str := 'Tropensturm';
			02:	str := 'Wirbelsturm';
			03:	str := 'starkes Gewitter ';
			04:	str := 'Gewitter';
			05:	str := 'Schneeregen';
			06:	str := 'Schneeregen';
			07:	str := 'Schneeregen';
			08:	str := 'gefrierender Nieselregen';
			09:	str := 'Nieselregen';
			10:	str := 'gefrierender Regen';
			11:	str := 'sertsehn';
			12:	str := 'sertstrets';
			13:	str := 'sjstj';
			14:	str := 'leichte yrderew';
			15:	str := 'Schneetreiben';
			16:	str := 'Schnee';
			17:	str := 'Hagel';
			18:	str := 'Schneeregen';
			19:	str := 'Staub';
			20:	str := 'nebelig';
			21:	str := 'Dunst';
			22:	str := 'rauchig';
			23:	str := 'sertsert';
			24:	str := 'windig';
			25:	str := 'kalt';
			26:	str := 'sertsert';
			27:	str := 'meist sertsert';
			28:	str := 'meist sertsert';
			29:	str := 'teilweise serhser';
			30:	str := 'teilweise sertsertshe';
			31:	str := 'klar';
			32:	str := 'sonnig';
			33:	str := 'heiter';
			34:	str := 'heiter';
			35:	str := 'Regen und Hagel';
			36:	str := 'WRYTWRYH';
			37:	str := 'esrertsertr';
			38:	str := 'vereinzelte Gewitter';
			39:	str := 'vereinzelte Gewitter';
			40:	str := 'verteesr';
			41:	str := 'sjstjtj';
			42:	str := 'sertsert';
			43:	str := 'sertsert';
			44:	str := 'sertsert';
			45:	str := 'sertsert';
			46:	str := 'sertsert';
			47:	str := 'srtsert';
			ELSE
				str := 'sertsert';
			END_CASE;
		END_FOR;
	END_IF;
	act_last := ACTIVATE;

END_FUNCTION_BLOCK

PROGRAM program0
	VAR
		ACTIVATE :	BOOL;
		YW :	oscat_YAHOO_WEATHER_DATA;

		func_block : YAHOO_WEATHER_DESC_GE_Block;
	END_VAR
	func_block.ACTIVATE := ACTIVATE;
	func_block.YW := YW;

	func_block();
	YW  := func_block.YW;
END_PROGRAM

CONFIGURATION Config0
	RESOURCE Res0 ON PLC
		TASK task0(INTERVAL := T#20ms,PRIORITY := 0);
		PROGRAM instance0 WITH task0 : program0;
	END_RESOURCE
END_CONFIGURATION

(* ---- 738-OSCAT.IEC ---- *)
(*@PROPERTIES_EX@
TYPE: DATA_TYPE
LOCALE: 0
*)
TYPE
  oscat_STRING1               : STRING(1);
  oscat_STRING2               : STRING(2);
  oscat_STRING3               : STRING(3);
  oscat_STRING4               : STRING(4);
  oscat_STRING5               : STRING(5);
  oscat_STRING8               : STRING(8);
  oscat_STRING10              : STRING(10);
  oscat_STRING12              : STRING(12);
  oscat_STRING15              : STRING(15);
  oscat_STRING20              : STRING(20);
  oscat_STRING27              : STRING(27);
  oscat_STRING30              : STRING(30);
  oscat_STRING32              : STRING(32);
  oscat_STRING40              : STRING(40);
  oscat_STRING48              : STRING(48);
  oscat_STRING50              : STRING(50);
  oscat_STRING60              : STRING(60);
  oscat_STRING64              : STRING(64);
  oscat_STRING80              : STRING(80);
  oscat_STRING120             : STRING(120);
  oscat_STRING144             : STRING(144);
  oscat_STRING160             : STRING(160);
  oscat_STRING189             : STRING(189);
  oscat_STRING192             : STRING(192);
  oscat_STRING250             : STRING(250);
END_TYPE

(*----------------------------------------------------------------------------------*)
TYPE

  oscat_arr_0_7               : ARRAY [0..7]    OF REAL;
  oscat_arr_0_15              : ARRAY [0..15]   OF REAL;
  oscat_delay_buf             : ARRAY [0..31]   OF REAL;
  oscat_FT_TN64_array         : ARRAY [0..63]   OF REAL;
  oscat_pt_ARRAY              : ARRAY [1..100]  OF REAL;

  oscat_ardw_0_15             : ARRAY [0..15]   OF DWORD;
  oscat_ardw_0_31             : ARRAY [0..31]   OF DWORD;

  oscat_FILTER_MAV_W          : ARRAY [0..31]   OF WORD;
  oscat_arb_0_3               : ARRAY [0..3]    OF BYTE;

  oscat_esr_collect_data      : ARRAY [0..7]    OF BYTE;
  oscat_DRIVER_4C 			  : ARRAY [1..7] 	OF BYTE;
  oscat_arb_0_249 			  : ARRAY [0..249] 	OF BYTE;
  oscat_bya_LIST_CLEAN        : ARRAY [1..250]  OF BYTE;

  oscat_ari_0_30         	  : ARRAY [0..30]   OF INT;

  oscat_stack_array 		  : ARRAY [1..32]   OF INT;

  oscat_dcf77_bits            : ARRAY [0..58]   OF BOOL;

  oscat_array64_time          : ARRAY [0..63]   OF TIME;

  (* -------------------------------------------------- *)
  oscat_PERIOD2_Y             : ARRAY [0..1]    OF UDINT;
  oscat_PERIOD2_X             : ARRAY [0..3]    OF oscat_PERIOD2_Y;

  oscat_ARRAY_X               : ARRAY [0..1]    OF REAL;
  oscat_XY                    : ARRAY [1..20]   OF oscat_ARRAY_X;

  oscat_parset_X              : ARRAY [1..4]    OF REAL;
  oscat_parset                : ARRAY [0..3]    OF oscat_parset_X;

  oscat_Polynom_ARRAY_X       : ARRAY [0..1]    OF REAL;
  oscat_Polynom_XY            : ARRAY [1..5]    OF oscat_Polynom_ARRAY_X;

END_TYPE

(*----------------------------------------------------------------------------------*)
TYPE oscat_FRACTION :
STRUCT
	NUMERATOR : INT;
	DENOMINATOR : INT;
END_STRUCT;
END_TYPE
(*----------------------------------------------------------------------------------*)
TYPE oscat_CALENDAR :
	STRUCT
		UTC : UDINT;				(* world time UTC *)
		LDT : UDINT;				(* local time *)
		LDATE : UDINT;				(* local date *)
		LTOD : UDINT;				(* local time of day *)
		YEAR : INT;					(* year of LDATE *)
		MONTH : INT;				(* month of LDATE *)
		DAY : INT;					(* day of LDATE *)
		WEEKDAY : INT;				(* weekday of LDATE *)
		OFFSET : INT;				(* Time Zone Offset for Local time in minutes *)
		DST_EN : BOOL;				(* daylight savings time enable *)
		DST_ON : BOOL;				(* true when daylight savings time os on *)
		NAME : oscat_string5;		(* name of time zone *)
		LANGUAGE : INT;			    (* language number pls see language setup *)
		LONGITUDE : REAL;			(* longitude of current location *)
		LATITUDE : REAL;			(* latitude of current location *)
		SUN_RISE : UDINT;			(* sun_rise for current location *)
		SUN_SET : UDINT;			(* sun_set for current location *)
		SUN_MIDDAY : UDINT;			(* worldtime when sun stands at south position *)
		SUN_HEIGTH : REAL;			(* suns heigth at midday, south position *)
		SUN_HOR : REAL;				(* sun angle horizontal 0 = north in degrees *)
		SUN_VER : REAL;				(* sun angle vertical above horizon in degrees *)
		NIGHT : BOOL;				(* true between sun_set and sun_rise *)
		HOLIDAY : BOOL;				(* true when holiday *)
		HOLY_NAME : oscat_string30;	(* name of holiday *)
		WORK_WEEK : INT;			(* current work week *)
	END_STRUCT;
END_TYPE

TYPE oscat_SDT :
STRUCT
	YEAR : INT;
	MONTH : INT;
	DAY : INT;
	WEEKDAY : INT;
	HOUR : INT;
	MINUTE : INT;
	SECOND : INT;
	MS : INT;
END_STRUCT;
END_TYPE

(*----------------------------------------------------------------------------------*)

TYPE oscat_LANGUAGE:
  STRUCT
    DEFAULT 	: INT;
	LMAX    	: INT;
  END_STRUCT;
END_TYPE

(*----------------------------------------------------------------------------------*)
TYPE
	oscat_LOCATION_ELEMENTS	: ARRAY [1..5] OF INT;
END_TYPE

TYPE oscat_LOCATION:
  STRUCT
    DEFAULT 	: INT;
	LMAX    	: INT;
	LANGUAGE	: oscat_LOCATION_ELEMENTS;
  END_STRUCT;
END_TYPE

(*----------------------------------------------------------------------------------*)

TYPE
  oscat_ELEMENT_DIRS 		: ARRAY [0..15] OF oscat_STRING3;
  oscat_DIRS				: ARRAY [1..3]  OF oscat_ELEMENT_DIRS;
END_TYPE

(*----------------------------------------------------------------------------------*)
TYPE
  oscat_CHARNAMES	: ARRAY [1..11] OF STRING;
END_TYPE

(*----------------------------------------------------------------------------------*)

TYPE
  oscat_ELEMENT_MONTHS 	: ARRAY [1..12] OF oscat_STRING10;
  oscat_MONTHS			: ARRAY [1..3]  OF oscat_ELEMENT_MONTHS;
END_TYPE

(*----------------------------------------------------------------------------------*)

TYPE
  oscat_ELEMENT_MONTHS3	: ARRAY [1..12] OF oscat_STRING3;
  oscat_MONTHS3			: ARRAY [1..3]  OF oscat_ELEMENT_MONTHS3;
END_TYPE

(*----------------------------------------------------------------------------------*)

TYPE
  oscat_ELEMENT_WEEKDAYS	: ARRAY [1..7] OF oscat_STRING10;
  oscat_WEEKDAYS			: ARRAY [1..3]  OF oscat_ELEMENT_WEEKDAYS;
END_TYPE

(*----------------------------------------------------------------------------------*)

TYPE
  oscat_ELEMENT_WEEKDAYS2	: ARRAY [1..7] OF oscat_STRING2;
  oscat_WEEKDAYS2			: ARRAY [1..3]  OF oscat_ELEMENT_WEEKDAYS2;
END_TYPE

TYPE oscat_esr_data :
  STRUCT
	typ    : BYTE;
	adress : oscat_string10;
	DS     : UDINT;
	TS     : TIME;
	data   : oscat_esr_collect_data;
  END_STRUCT;
END_TYPE

TYPE
  oscat_ESR_3                : ARRAY [0..3] OF oscat_esr_data;
  oscat_ESR_31               : ARRAY [0..31] OF oscat_esr_data;
END_TYPE

TYPE oscat_vector_3 :
  STRUCT
	X : REAL;
	Y : REAL;
	Z : REAL;
  END_STRUCT;
END_TYPE

TYPE oscat_complex :
  STRUCT
	re : REAL;
	im : REAL;
  END_STRUCT;
END_TYPE

TYPE REAL2 :
  STRUCT
	R1 : REAL;
	RX : REAL;
  END_STRUCT;
END_TYPE

(*----------------------------------------------------------------------------------*)

TYPE oscat_HOLIDAY_DATA :
  STRUCT
	NAME : oscat_string30;
	DAY : SINT;
	MONTH : SINT;
	USE : SINT;
	PAD_BYTE : BYTE;
  END_STRUCT;
END_TYPE

TYPE
  oscat_HOLIDAY_DATA_0_29 	: ARRAY [0..29] OF oscat_HOLIDAY_DATA;
  oscat_HOLIDAY_DATA_0_49 	: ARRAY [0..49] OF oscat_HOLIDAY_DATA;
END_TYPE

(* revision history
hm	18. oct. 2008
	original version

*)

(*	if month = 0 then F_day is the offset in days from easter
	used :0 = NOT used, 1 = used, -1..-7 menas the weekday before the specified DATE example -3 means wednesday before 23.11
*)

(* samples for Holiday data

	HOLIDAY_DE : ARRAY[0..29] OF HOLIDAY_DATA := (name := 'Neujahr', day := 1, month := 1, use := 1),
		(name := 'Heilig Drei Könige', day := 6, month := 1, use := 1),
		(name := 'Karfreitag', day := -2, month := 0, use := 1),
		(name := 'Ostersonntag', day := 0, month := 0, use := 1),
		(name := 'Ostermontag', day := 1, month := 0, use := 1),
		(name := 'Tag der Arbeit', day := 1, month := 5, use := 1),
		(name := 'Christi Himmelfahrt', day := 39, month := 0, use := 1),
		(name := 'Pfingstsonntag', day := 49, month := 0, use := 1),
		(name := 'Pfingstmontag', day := 50, month := 0, use := 1),
		(name := 'Fronleichnam', day := 60, month := 0, use := 1),
		(name := 'Augsburger Friedensfest', day := 8, month := 8, use := 0),
		(name := 'Maria Himmelfahrt', day := 15, month := 8, use := 1),
		(name := 'Tag der Deutschen Einheit', day := 3, month := 10, use := 1),
		(name := 'Reformationstag', day := 31, month := 10, use := 0),
		(name := 'Allerheiligen', day := 1, month := 11, use := 1),
		(name := 'Buss und Bettag', day := 23, month := 11, use := 0),
		(name := '1. Weihnachtstag', day := 25, month := 12, use := 1),
		(name := '2. Weihnachtstag', day := 26, month := 12, use := 1);

	HOLIDAY_AT : ARRAY[0..29] OF HOLIDAY_DATA := (name := 'Neujahr', day := 1, month := 1, use := 1),
		(name := 'Heilig Drei Könige', day := 6, month := 1, use := 1),
		(name := 'Karfreitag', day := -2, month := 0, use := 1),
		(name := 'Ostersonntag', day := 0, month := 0, use := 1),
		(name := 'Ostermontag', day := 1, month := 0, use := 1),
		(name := '', day := 1, month := 5, use := 0),
		(name := 'Christi Himmelfahrt', day := 39, month := 0, use := 1),
		(name := 'Pfingstsonntag', day := 49, month := 0, use := 1),
		(name := 'Pfingstmontag', day := 50, month := 0, use := 1),
		(name := 'Fronleichnam', day := 60, month := 0, use := 1),
		(name := '', day := 8, month := 8, use := 0),
		(name := 'Maria Himmelfahrt', day := 15, month := 8, use := 1),
		(name := '', day := 3, month := 10, use := 0),
		(name := '', day := 31, month := 10, use := 0),
		(name := 'Allerheiligen', day := 1, month := 11, use := 1),
		(name := 'Maria Empfängnis', day := 8, month := 12, use := 1),
		(name := '1. Weihnachtstag', day := 25, month := 12, use := 1),
		(name := '2. Weihnachtstag', day := 26, month := 12, use := 1);

	HOLIDAY_FR : ARRAY[0..29] OF HOLIDAY_DATA := (name := 'Nouvel an', day := 1, month := 1, use := 1),
		(name := 'St Valentin', day := 14, month := 2, use := 0),
		(name := 'Vendredi Saint (alsace)', day := -2, month := 0, use := 0),
		(name := 'Dimanche de pâques', day := 0, month := 0, use := 1),
		(name := 'Lundi de pâques', day := 1, month := 0, use := 1),
		(name := 'Jeudi de Ascension', day := 39, month := 0, use := 1),
		(name := 'dimanche de Pentecôte ', day := 49, month := 0, use := 1),
		(name := 'jeudi de la Trinité', day := 60, month := 0, use := 0),
		(name := 'Fête du travail', day := 1, month := 5, use := 1),
		(name := 'Victoire 1945 ', day := 8, month := 5, use := 1),
		(name := 'Prise de La bastille', day := 14, month := 7, use := 1),
		(name := '15 Août 1944', day := 15, month := 8, use := 1),
		(name := 'Halloween', day := 31, month := 10, use := 0),
		(name := 'Armistice 1918', day := 11, month := 11, use := 1),
		(name := 'Noël', day := 25, month := 12, use := 1),
		(name := 'Saint Étienne (alsace)', day := 26, month := 12, use := 0),
		(name := 'Fête de la musique', day := 21, month := 6, use := 0);

	HOLIDAY_BED : ARRAY[0..29] OF HOLIDAY_DATA :=	(name := 'Neujahr', day := 1, month := 1, use := 1),
		(name := 'Ostersonntag', day := 0, month := 0, use := 1),
		(name := 'Ostermontag', day := 1, month := 0, use := 1),
		(name := 'Tag der Arbeit', day := 1, month := 5, use := 1),
		(name := 'Christi Himmelfahrt', day := 39, month := 0, use := 1),
		(name := 'Pfingsten', day := 49, month := 0, use := 1),
		(name := 'Pfingstmontag', day := 50, month := 0, use := 1),
		(name := 'Nationalfeiertag', day := 21, month := 7, use := 1),
		(name := 'Mariä Himmelfahrt', day := 15, month := 8, use := 1),
		(name := 'Allerheiligen', day := 1, month := 11, use := 1),
		(name := 'Feiertag DG', day := 15, month := 11, use := 1),
		(name := 'Heiligabend', day := 24, month := 12, use := 1),
		(name := '1. Weihnachtstag', day := 25, month := 12, use := 1),
		(name := '2. Weihnachtstag', day := 26, month := 12, use := 1),
		(name := 'Silvester', day := 31, month := 12, use := 1);

	HOLIDAY_ITD : ARRAY[0..29] OF HOLIDAY_DATA := (name := 'Neujahr', day := 1, month := 1, use := 1),
		(name := 'Heilig Drei Könige', day := 6, month := 1, use := 1),
		(name := 'Ostersonntag', day := 0, month := 0, use := 1),
		(name := 'Ostermontag', day := 1, month := 0, use := 1),
		(name := 'Tag der Befeiung Italiens', day := 25, month := 4, use := 1),
		(name := 'Tag der Arbeit', day := 1, month := 5, use := 1),
		(name := 'Pfingsten', day := 49, month := 0, use := 1),
		(name := 'Pfingstmontag', day := 50, month := 0, use := 1),
		(name := 'Tag der Republik Italien', day := 2, month := 6, use := 1),
		(name := 'Mariä Himmelfahrt', day := 15, month := 8, use := 1),
		(name := 'Allerheiligen', day := 1, month := 11, use := 1),
		(name := 'Mariä Empfängnis', day := 8, month := 12, use := 1),
		(name := 'Heiligabend', day := 24, month := 12, use := 0),
		(name := '1. Weihnachtstag', day := 25, month := 12, use := 1),
		(name := '2. Stephanstag', day := 26, month := 12, use := 1);

*)

(* ---- 740-TIMER_P4.ST ---- *)
TYPE oscat_TIMER_EVENT_DATA :
  STRUCT
	TYP          : BYTE;
	CHANNEL      : BYTE;
	DAY          : BYTE;
	START        : UDINT;
	DURATION     : TIME;
	LAND         : BYTE;
	LOR          : BYTE;
	LAST         : UDINT;
  END_STRUCT;
END_TYPE

TYPE
  oscat_TIMER_EVENT           : ARRAY [0..63]    OF oscat_TIMER_EVENT_DATA;
  oscat_TP4_qn                : ARRAY [0..3]    OF BOOL;
END_TYPE

TYPE
  oscat_arb_0_3               : ARRAY [0..3]    OF BYTE;
END_TYPE

FUNCTION _BYTE_TO_INT:INT
	VAR_INPUT
		IN :	BYTE;
	END_VAR

	_BYTE_TO_INT := USINT_TO_INT(BYTE_TO_USINT(IN));
END_FUNCTION

FUNCTION DATE_TO_DT:UDINT
	VAR_INPUT
		IN :	UDINT;
	END_VAR
	DATE_TO_DT := IN;
END_FUNCTION

FUNCTION _DT_TO_DATE_B:UDINT

	VAR_INPUT
		_INN :	UDINT;
	END_VAR

	_DT_TO_DATE_B := (_INN / UDINT#86400) * UDINT#86400;
END_FUNCTION

FUNCTION TIME_TO_UDINT2:UDINT
	VAR_INPUT
		X :	TIME;
	END_VAR

	TIME_TO_UDINT2 := DINT_TO_UDINT(TIME_TO_DINT(X));
END_FUNCTION

FUNCTION DATE_TO_UDINT2:UDINT
	VAR_INPUT
		IN :	UDINT;
	END_VAR

	DATE_TO_UDINT2 := IN;
END_FUNCTION

FUNCTION DAY_OF_WEEK:INT
  VAR_INPUT
    IDATE :	UDINT;
  END_VAR

  DAY_OF_WEEK := UDINT_TO_INT((idate / UDINT#86400 + UDINT#3) MOD UDINT#7) + INT#01;
END_FUNCTION

FUNCTION _BYTE_TO_DINT:DINT
	VAR_INPUT
		IN :	BYTE;
	END_VAR

	_BYTE_TO_DINT := USINT_TO_DINT(BYTE_TO_USINT(IN));
END_FUNCTION

FUNCTION DAY_OF_YEAR_UDINT:INT
	VAR_INPUT
		IDATE :	UDINT;
	END_VAR

	DAY_OF_YEAR_UDINT := UDINT_TO_INT((idate / UDINT#86400) MOD UDINT#1461);
	IF DAY_OF_YEAR_UDINT > 729 THEN
		IF DAY_OF_YEAR_UDINT > 1095 THEN DAY_OF_YEAR_UDINT := DAY_OF_YEAR_UDINT - 1095; ELSE DAY_OF_YEAR_UDINT := DAY_OF_YEAR_UDINT - 729; END_IF;
	ELSIF DAY_OF_YEAR_UDINT > 364 THEN
		DAY_OF_YEAR_UDINT := DAY_OF_YEAR_UDINT - 364;
	ELSE
		DAY_OF_YEAR_UDINT := DAY_OF_YEAR_UDINT + 1;
	END_IF;
END_FUNCTION

FUNCTION MONTH_OF_DATE_UDINT:INT

	VAR_INPUT
		IDATE :	UDINT;
	END_VAR

	MONTH_OF_DATE_UDINT := DAY_OF_YEAR_UDINT(idate);
	IF MONTH_OF_DATE_UDINT < 32 THEN
		MONTH_OF_DATE_UDINT := 1;
	ELSIF LEAP_OF_DATE(IDATE) THEN
		MONTH_OF_DATE_UDINT := (MONTH_OF_DATE_UDINT * 53 + 1668) / 1623;
	ELSE
		MONTH_OF_DATE_UDINT := (MONTH_OF_DATE_UDINT * 53 + 1700) / 1620;
	END_IF;

END_FUNCTION

FUNCTION DAY_OF_MONTH:INT
	VAR_INPUT
		IDATE :	UDINT;
	END_VAR

	day_of_month := day_of_year_UDINT(idate);

	IF leap_of_Date(idate) THEN
		CASE day_of_month OF
			32..60	:	day_of_month := day_of_month - 31;
			61..91	:	day_of_month := day_of_month - 60;
			92..121 :	day_of_month := day_of_month - 91;
			122..152:	day_of_month := day_of_month - 121;
			153..182:	day_of_month := day_of_month - 152;
			183..213:	day_of_month := day_of_month - 182;
			214..244:	day_of_month := day_of_month - 213;
			245..274:	day_of_month := day_of_month - 244;
			275..305:	day_of_month := day_of_month - 274;
			306..335:	day_of_month := day_of_month - 305;
			336..366:	day_of_month := day_of_month - 335;
		END_CASE;
	ELSE
		CASE day_of_month OF
			32..59	:	day_of_month := day_of_month - 31;
			60..90	:	day_of_month := day_of_month - 59;
			91..120 :	day_of_month := day_of_month - 90;
			121..151:	day_of_month := day_of_month - 120;
			152..181:	day_of_month := day_of_month - 151;
			182..212:	day_of_month := day_of_month - 181;
			213..243:	day_of_month := day_of_month - 212;
			244..273:	day_of_month := day_of_month - 243;
			274..304:	day_of_month := day_of_month - 273;
			305..334:	day_of_month := day_of_month - 304;
			335..365:	day_of_month := day_of_month - 334;
		END_CASE;
	END_IF;

END_FUNCTION

FUNCTION LEAP_OF_DATE:BOOL

	VAR_INPUT
		IDATE :	UDINT;
	END_VAR

	LEAP_OF_DATE := SHL(UDINT_TO_DWORD((idate + UDINT#43200) / UDINT#31557600), 30) = DWORD#16#80000000;
END_FUNCTION

FUNCTION DAY_OF_YEAR:INT
	VAR_INPUT
		IDATE :	UDINT;
	END_VAR

	DAY_OF_YEAR := UDINT_TO_INT(((idate) / UDINT#86400) MOD UDINT#1461);
	IF DAY_OF_YEAR > 729 THEN
		IF DAY_OF_YEAR > 1095 THEN DAY_OF_YEAR := DAY_OF_YEAR - 1095; ELSE DAY_OF_YEAR := DAY_OF_YEAR - 729; END_IF;
	ELSIF DAY_OF_YEAR > 364 THEN
		DAY_OF_YEAR := DAY_OF_YEAR - 364;
	ELSE
		DAY_OF_YEAR := DAY_OF_YEAR + 1;
	END_IF;
END_FUNCTION

FUNCTION MONTH_OF_DATE:INT

	VAR_INPUT
		IDATE :	UDINT;
	END_VAR

	MONTH_OF_DATE := DAY_OF_YEAR(idate);
	IF MONTH_OF_DATE < 32 THEN
		MONTH_OF_DATE := 1;
	ELSIF LEAP_OF_DATE((IDATE)) THEN
		MONTH_OF_DATE := (MONTH_OF_DATE * 53 + 1668) / 1623;
	ELSE
		MONTH_OF_DATE := (MONTH_OF_DATE * 53 + 1700) / 1620;
	END_IF;
END_FUNCTION

FUNCTION YEAR_OF_DATE:INT
	VAR_INPUT
		IDATE :	UDINT;
	END_VAR

	YEAR_OF_DATE := UDINT_TO_INT((idate+UDINT#43200) / UDINT#31557600 + UDINT#1970);
END_FUNCTION

FUNCTION _INT_TO_UDINT:UDINT
	VAR_INPUT
		IN :	INT;
	END_VAR

	_INT_TO_UDINT := DINT_TO_UDINT(INT_TO_DINT(IN));
END_FUNCTION

FUNCTION DT_TO_DATE:UDINT
	VAR_INPUT
		IN :	UDINT;
	END_VAR

	DT_TO_DATE := (IN / UDINT#86400) * UDINT#86400;
END_FUNCTION

FUNCTION SET_DT:UDINT

	VAR_INPUT
		YEAR : INT;
		MONTH :	INT;
		DAY : INT;
		HOUR : INT;
		MINUTE : INT;
		SECOND : INT;
	END_VAR

	SET_DT := SET_DATE(YEAR, MONTH, DAY) + _INT_TO_UDINT(SECOND) + _INT_TO_UDINT(MINUTE) * UDINT#60 + _INT_TO_UDINT(HOUR) * UDINT#3600;

END_FUNCTION

FUNCTION SET_DATE:UDINT

	VAR_INPUT
		YEAR :	INT;
		MONTH :	INT;
		DAY :	INT;
	END_VAR

	VAR
		count :	INT;
	END_VAR

	IF month > 2 THEN
		count := (month - 1) * 30;
		IF month > 7 THEN
			count := count + DWORD_TO_INT(SHR(DINT_TO_DWORD(INT_TO_DINT(month) - INT_TO_DINT(3)),1));
		ELSE
			count := count + DWORD_TO_INT(SHR(DINT_TO_DWORD(INT_TO_DINT(month) - INT_TO_DINT(4)),1));
		END_IF;
		IF SHL(INT_TO_WORD(year),14) = WORD#0 THEN
			count := count + 1;
		END_IF;
	ELSE
		count := (month - 1) * 31;
	END_IF;
	SET_DATE := (_INT_TO_UDINT(count + day - 1) + DWORD_TO_UDINT(SHR(UDINT_TO_DWORD(_INT_TO_UDINT(year) * UDINT#1461 - UDINT#2878169), 2))) * UDINT#86400;

END_FUNCTION

FUNCTION MONTH_END:UDINT

	VAR_INPUT
		IDATE :	UDINT;
	END_VAR

	MONTH_END := SET_DATE(YEAR_OF_DATE(idate),MONTH_OF_DATE(idate)+1,1) - UDINT#86400;

END_FUNCTION

FUNCTION YEAR_END:UDINT

	VAR_INPUT
		Y :	INT;
	END_VAR

	YEAR_END := DWORD_TO_UDINT(SHR(UDINT_TO_DWORD(INT_TO_UDINT(y) * UDINT#1461 - UDINT#2876712), 2)) * UDINT#86400;

END_FUNCTION

FUNCTION LEAP_DAY:BOOL

	VAR_INPUT
		IDATE :	UDINT;
	END_VAR

	LEAP_DAY := IDATE MOD UDINT#126230400 = UDINT#68169600;

END_FUNCTION

FUNCTION BIT_LOAD_B:BYTE
	VAR_INPUT
		IN :	BYTE;
		VAL :	BOOL;
		POS :	INT;
	END_VAR

	IF VAL THEN
		BIT_LOAD_B := in OR SHL(BYTE#1,pos);
	ELSE
		BIT_LOAD_B := in AND (NOT SHL(BYTE#1,pos));
	END_IF;
END_FUNCTION

FUNCTION BIT_OF_DWORD : BOOL
  VAR_INPUT
    IN : DWORD;
    N : INT;
  END_VAR

  BIT_OF_DWORD := (SHR(in,N) AND 16#00000001) > 0;
END_FUNCTION

FUNCTION_BLOCK TIMER_P4_Block

	VAR_INPUT
		DTIME :	UDINT;
		TREF_0 :	UDINT;
		TREF_1 :	UDINT;
		HOLY :	BOOL;
		L0 :	BOOL;
		L1 :	BOOL;
		L2 :	BOOL;
		L3 :	BOOL;
		OFS :	BYTE;
		ENQ :	BOOL;
		MAN :	BOOL;
		MI :	BYTE;
		RST :	BOOL;
	END_VAR

	VAR_IN_OUT
		PROG :	oscat_TIMER_EVENT;
	END_VAR

	VAR_OUTPUT
		Q0 :	BOOL;
		Q1 :	BOOL;
		Q2 :	BOOL;
		Q3 :	BOOL;
		STATUS :	BYTE;
	END_VAR

	VAR
		day_start :	UDINT;
		start :	UDINT;
		event :	oscat_TIMER_EVENT_DATA;
		pos :	INT;
		last_execute :	UDINT;
		current_day :	DINT;
		mask :	BYTE;
		ma :	oscat_arb_0_3;
		mo :	oscat_arb_0_3;
		qn :	oscat_TP4_qn;
		qs :	oscat_TP4_qn;
		channel :	INT;
		tx :	UDINT;
		array_max :	INT := 63;
		channel_max :	INT := 3;
	END_VAR

	IF RST THEN
		last_execute := UDINT#00;
		FOR pos := 0 TO ARRAY_MAX DO
			IF (PROG[pos].CHANNEL >= OFS) AND (_BYTE_TO_INT(PROG[pos].CHANNEL) < (_BYTE_TO_INT(OFS) + 4)) THEN PROG[pos].LAST := last_execute; END_IF;
		END_FOR;

		FOR pos := 0 TO channel_max DO
			qs[pos] := FALSE;
		END_FOR;

	ELSIF dtime <> last_execute THEN
		last_execute := DTIME;

		day_start := DATE_TO_DT(_DT_TO_DATE_B(DTIME));

		FOR pos := 0 TO channel_max DO qn[pos] := FALSE; END_FOR;

		FOR pos := 0 TO ARRAY_MAX DO
			event := prog[pos];
			channel := _BYTE_TO_INT(event.CHANNEL) - _BYTE_TO_INT(OFS);
			IF (event.TYP > BYTE#0) AND (channel >= 0) AND (channel <= channel_max) THEN
				ma[channel] := event.LAND;
				mo[channel] := event.LOR;
				CASE _BYTE_TO_INT(event.TYP) OF
					1:
						start := day_start + event.start;
						qn[channel] := dtime >= start AND dtime <= start + TIME_TO_UDINT2(event.DURATION);

					2:
						IF (SHR(BYTE#128, DAY_OF_WEEK(_DT_TO_DATE_B(Dtime))) AND event.DAY) > BYTE#0 THEN
							start := day_start + event.start;
							qn[channel] := dtime >= start AND dtime <= start + TIME_TO_UDINT2(event.DURATION);
						END_IF;

					3:
						IF current_day MOD _BYTE_TO_DINT(event.DAY) = DINT#0 THEN
							start := day_start + event.start;
							qn[channel] := dtime >= start AND dtime <= start + TIME_TO_UDINT2(event.DURATION);
						END_IF;

					10:
						IF DAY_OF_WEEK(_DT_TO_DATE_B(DTIME)) = BYTE_TO_INT(event.DAY) THEN
							start := day_start + event.start;
							qn[channel] := dtime >= start AND dtime <= start + TIME_TO_UDINT2(event.DURATION);
						END_IF;

					20:
						IF DAY_OF_MONTH(_DT_TO_DATE_B(DTIME)) = BYTE_TO_INT(event.DAY) THEN
							start := day_start + event.start;
							qn[channel] := dtime >= start AND dtime <= start + TIME_TO_UDINT2(event.DURATION);
						END_IF;

					21:
						IF _DT_TO_DATE_B(DTIME) = MONTH_END(_DT_TO_DATE_B(dtime)) THEN
							start := day_start + event.start;
							qn[channel] := dtime >= start AND dtime <= start + TIME_TO_UDINT2(event.DURATION);
						END_IF;

					30:
						IF DAY_OF_YEAR(_DT_TO_DATE_B(DTIME)) = BYTE_TO_INT(event.DAY) THEN
							start := day_start + event.start;
							qn[channel] := dtime >= start AND dtime <= start + TIME_TO_UDINT2(event.DURATION);
						END_IF;

					31:
						IF _DT_TO_DATE_B(DTIME) = YEAR_END(YEAR_OF_DATE(_DT_TO_DATE_B(dtime))) THEN
							start := day_start + event.start;
							qn[channel] := dtime >= start AND dtime <= start + TIME_TO_UDINT2(event.DURATION);
						END_IF;

					40:
						IF LEAP_DAY(_DT_TO_DATE_B(dtime)) THEN
							start := day_start + event.start;
							qn[channel] := dtime >= start AND dtime <= start + TIME_TO_UDINT2(event.DURATION);
						END_IF;

					41:
						IF HOLY THEN
							start := day_start + event.start;
							qn[channel] := dtime >= start AND dtime <= start + TIME_TO_UDINT2(event.DURATION);
						END_IF;

					42:
						IF (Holy OR (DAY_OF_WEEK(_DT_TO_DATE_B(dtime)) = 6) OR (DAY_OF_WEEK(_DT_TO_DATE_B(dtime)) = 7)) THEN
							start := day_start + event.start;
							qn[channel] := dtime >= start AND dtime <= start + TIME_TO_UDINT2(event.DURATION);
						END_IF;

					43:
						IF DAY_OF_WEEK(_DT_TO_DATE_B(dtime)) < 6 THEN
							start := day_start + event.start;
							qn[channel] := dtime >= start AND dtime <= start + TIME_TO_UDINT2(event.DURATION);
						END_IF;

					50:
						CASE _BYTE_TO_INT(prog[pos].DAY) OF
							0:	tx := tref_0;
							1:	tx := tref_1;
						ELSE
							tx := UDINT#0 ;
						END_CASE;
						start := day_start + tx + event.start;
						qn[channel] := dtime >= start AND dtime <= start + TIME_TO_UDINT2(event.DURATION);

					51:
						CASE _BYTE_TO_INT(prog[pos].DAY) OF
							0:	tx := tref_0;
							1:	tx := tref_1;
						ELSE
							tx := UDINT#0;
						END_CASE;
						start := day_start + tx - event.start;
						qn[channel] := dtime >= start AND dtime <= start + TIME_TO_UDINT2(event.DURATION);

					52 :
						CASE _BYTE_TO_INT(prog[pos].DAY) OF
							0:	tx := tref_0;
							1:	tx := tref_1;
						ELSE
							tx := UDINT#0 ;
						END_CASE;
						start := day_start + tx + event.start;
						IF dtime >= start AND day_start > event.LAST THEN
							qs[channel] := TRUE;
							prog[pos].LAST := day_start;
						END_IF;

					53 :
						CASE _BYTE_TO_INT(prog[pos].DAY) OF
							0:	tx := tref_0;
							1:	tx := tref_1;
						ELSE
							tx := UDINT#0 ;
						END_CASE;
						start := day_start + tx + event.start;
						IF dtime >= start AND day_start > event.LAST THEN
							qs[channel] := FALSE;
							prog[pos].LAST := day_start;
						END_IF;

					54 :
						CASE _BYTE_TO_INT(prog[pos].DAY) OF
							0:	tx := tref_0;
							1:	tx := tref_1;
						ELSE
							tx := UDINT#0 ;
						END_CASE;
						start := day_start + tx - event.start;
						IF dtime >= start AND day_start > event.LAST THEN
							qs[channel] := TRUE;
							prog[pos].LAST := day_start;
						END_IF;

					55 :
						CASE _BYTE_TO_INT(prog[pos].DAY) OF
							0:	tx := tref_0;
							1:	tx := tref_1;
						ELSE
							tx := UDINT#0 ;
						END_CASE;
						start := day_start + tx - event.start;
						IF dtime >= start AND day_start > event.LAST THEN
							qs[channel] := FALSE;
							prog[pos].LAST := day_start;
						END_IF;
				END_CASE;
			END_IF;
		END_FOR;
	END_IF;

	mask := BYTE#255;
	mask:=BIT_LOAD_B(mask,L0,0);
	mask:=BIT_LOAD_B(mask,L1,1);
	mask:=BIT_LOAD_B(mask,L2,2);
	mask:=BIT_LOAD_B(mask,L3,3);

	Q0 := ENQ AND ((qn[0] OR qs[0]) AND ((ma[0] AND mask) = ma[0]) OR ((mo[0] AND mask) > BYTE#0) OR (man AND BIT_OF_DWORD(BYTE_TO_DWORD(MI),0)));
	Q1 := ENQ AND ((qn[1] OR qs[1]) AND ((ma[1] AND mask) = ma[1]) OR ((mo[1] AND mask) > BYTE#1) OR (man AND BIT_OF_DWORD(BYTE_TO_DWORD(MI),1)));
	Q2 := ENQ AND ((qn[2] OR qs[2]) AND ((ma[2] AND mask) = ma[2]) OR ((mo[2] AND mask) > BYTE#2) OR (man AND BIT_OF_DWORD(BYTE_TO_DWORD(MI),2)));
	Q3 := ENQ AND ((qn[3] OR qs[3]) AND ((ma[3] AND mask) = ma[3]) OR ((mo[3] AND mask) > BYTE#3) OR (man AND BIT_OF_DWORD(BYTE_TO_DWORD(MI),3)));

	IF NOT enq THEN
		status := BYTE#100;
	ELSIF man THEN
		status := BYTE#101;
	ELSE
		status := BYTE#102;
	END_IF;

END_FUNCTION_BLOCK

PROGRAM program0
	VAR
		DTIME :	UDINT;
		TREF_0 :	UDINT;
		TREF_1 :	UDINT;
		HOLY :	BOOL;
		L0 :	BOOL;
		L1 :	BOOL;
		L2 :	BOOL;
		L3 :	BOOL;
		OFS :	BYTE;
		ENQ :	BOOL;
		MAN :	BOOL;
		MI :	BYTE;
		RST :	BOOL;
		PROG :	oscat_TIMER_EVENT;
		Q0 :	BOOL;
		Q1 :	BOOL;
		Q2 :	BOOL;
		Q3 :	BOOL;
		STATUS :	BYTE;

		func_block : TIMER_P4_Block;
	END_VAR
	func_block.DTIME := DTIME;
	func_block.TREF_0 := TREF_0;
	func_block.TREF_1 := TREF_1;
	func_block.HOLY := HOLY;
	func_block.L0 := L0;
	func_block.L1 := L1;
	func_block.L2 := L2;
	func_block.L3 := L3;
	func_block.OFS := OFS;
	func_block.ENQ := ENQ;
	func_block.MAN := MAN;
	func_block.MI := MI;
	func_block.RST := RST;
	func_block.PROG := PROG;

	func_block();
	PROG  := func_block.PROG;
	Q0  := func_block.Q0;
	Q1  := func_block.Q1;
	Q2  := func_block.Q2;
	Q3  := func_block.Q3;
	STATUS  := func_block.STATUS;
END_PROGRAM

CONFIGURATION Config0
	RESOURCE Res0 ON PLC
		TASK task0(INTERVAL := T#20ms,PRIORITY := 0);
		PROGRAM instance0 WITH task0 : program0;
	END_RESOURCE
END_CONFIGURATION

(* ---- 1-IS_IP4.ST ---- *)
FUNCTION_BLOCK IS_IP4

	VAR_INPUT
		STR :	STRING;
	END_VAR

	VAR_OUTPUT
		IS_IP4 :	BOOL;
	END_VAR

	VAR
		COUNT_CHAR :	COUNT_CHAR;
	END_VAR

	COUNT_CHAR(STR:=str,CHR:=BYTE#46);
	IS_IP4 := COUNT_CHAR.COUNT_CHAR = 3;

END_FUNCTION_BLOCK

(* ---- 121-DEC_TO_INT.ST ---- *)
FUNCTION_BLOCK DEC_TO_INT
	VAR_INPUT
		DEC :		STRING;
	END_VAR

	VAR_OUTPUT
		DEC_TO_INT :	INT;
	END_VAR

	VAR
		i :	INT;
		X :	INT;
		sign :	BOOL;
		stop :	INT;
	END_VAR

	DEC_TO_INT := 0;
	sign := FALSE;
	stop := LEN(dec);
	FOR I := 1 TO stop DO
		X := GET_CHAR(DEC,I);
		IF X > 47 AND X < 58 THEN
			DEC_TO_INT := DEC_TO_INT * 10 + X - 48;
		ELSIF X = 45 AND DEC_TO_INT = 0 THEN
			sign := TRUE;
		END_IF;
	END_FOR;
	IF sign THEN DEC_TO_INT := -DEC_TO_INT; END_IF;

END_FUNCTION_BLOCK

(* ---- 141-SH_T.ST ---- *)
FUNCTION_BLOCK SH_T_Block

	VAR_INPUT
		IN :	REAL;
		E :	BOOL;
	END_VAR

	VAR_OUTPUT
		OUT :	REAL;
	END_VAR

	IF E THEN out := in; END_IF;

END_FUNCTION_BLOCK

PROGRAM program0

	VAR
		IN :	REAL;
		E :	BOOL;
		OUT :	REAL;
		func_block : SH_T_Block;
	END_VAR
	func_block.IN  :=IN;
	func_block.E  :=E;
	func_block();
	OUT := func_block.OUT;

END_PROGRAM

CONFIGURATION Config0

	RESOURCE Res0 ON PLC
		TASK task0(INTERVAL := T#20ms,PRIORITY := 0);
		PROGRAM instance0 WITH task0 : program0;
	END_RESOURCE

END_CONFIGURATION

(* ---- 149-DW_TO_REAL.ST ---- *)
FUNCTION_BLOCK DW_TO_REAL_Block
  VAR_INPUT
    X :	DWORD;
  END_VAR

  VAR_OUTPUT
    DW_TO_REAL :	REAL;
  END_VAR

  VAR
    BUF_TO_REAL :	BUF_TO_REAL;
    i :	INT;
  END_VAR

  FOR I := 0 TO 1 DO
    BUF_TO_REAL.REQ        := I > 0;
    BUF_TO_REAL.BUF_FORMAT := FALSE;
    BUF_TO_REAL.BUF_OFFS   := DINT#0;
    BUF_TO_REAL.BUF_CNT    := DINT#4;
    BUF_TO_REAL.BUFFER     := X;
    BUF_TO_REAL.DST        := DW_TO_REAL;
    BUF_TO_REAL();
    X           := BUF_TO_REAL.BUFFER;
    DW_TO_REAL  := BUF_TO_REAL.DST;
  END_FOR;
END_FUNCTION_BLOCK

(* ---- 151-B_TRIG.ST ---- *)
FUNCTION_BLOCK B_TRIG
	VAR_INPUT
		CLK :	BOOL;
	END_VAR

	VAR_OUTPUT
		Q :	BOOL := FALSE;
	END_VAR

	VAR
		edge :	BOOL := FALSE;
	END_VAR

	Q := clk XOR edge;
	edge := CLK;
END_FUNCTION_BLOCK

PROGRAM program0
  VAR
    LocalVar0 : BOOL;
	LocalOUT  : BOOL;
	func_block : B_TRIG;
  END_VAR
	func_block.CLK := LocalVar0;
	func_block();
	LocalOUT := func_block.Q;

END_PROGRAM

CONFIGURATION Config0
  RESOURCE Res0 ON PLC
    TASK task0(INTERVAL := T#20ms,PRIORITY := 0);
    PROGRAM instance0 WITH task0 : program0;
  END_RESOURCE
END_CONFIGURATION

(* ---- 152-BYTE_TO_STRH.ST ---- *)
FUNCTION_BLOCK BYTE_TO_STRH_Block
	VAR_INPUT
		IN :	BYTE;
	END_VAR

	VAR_OUTPUT
		BYTE_TO_STRH :	STRING;
	END_VAR

	BYTE_TO_STRH:=BYTE_TO_STRING(IN);

END_FUNCTION_BLOCK

PROGRAM program0
  VAR
    LocalVar0 : BYTE;
	LocalOUT  : STRING;
	func_block : BYTE_TO_STRH_Block;
  END_VAR
	func_block.IN  := LocalVar0;
	func_block();
	LocalOUT := func_block.BYTE_TO_STRH;

END_PROGRAM

CONFIGURATION Config0
  RESOURCE Res0 ON PLC
    TASK task0(INTERVAL := T#20ms,PRIORITY := 0);
    PROGRAM instance0 WITH task0 : program0;
  END_RESOURCE
END_CONFIGURATION

(* ---- 156-CHR_TO_STRING.ST ---- *)
FUNCTION_BLOCK CHR_TO_STRING_Block
	VAR_INPUT
		C :	BYTE;
	END_VAR

	VAR_OUTPUT
		CHR_TO_STRING :	STRING;
	END_VAR

	CHR_TO_STRING := BYTE_TO_STRING(C);

END_FUNCTION_BLOCK

PROGRAM program0
  VAR
    LocalVar0 : BYTE;
	LocalOUT  : STRING;
	func_block : CHR_TO_STRING_Block;
  END_VAR
	func_block.C  := LocalVar0;
	func_block();
	LocalOUT := func_block.CHR_TO_STRING;
END_PROGRAM

CONFIGURATION Config0
  RESOURCE Res0 ON PLC
    TASK task0(INTERVAL := T#20ms,PRIORITY := 0);
    PROGRAM instance0 WITH task0 : program0;
  END_RESOURCE
END_CONFIGURATION

(* ---- 158-TMIN.ST ---- *)
FUNCTION_BLOCK TMIN

	VAR_INPUT
		IN :	BOOL;
		PT :	TIME;
	END_VAR

	VAR_OUTPUT
		Q :	BOOL;
	END_VAR

	VAR
		pm :	TP;
	END_VAR

	pm(in := IN, PT := PT);
	Q := IN OR pm.Q;

END_FUNCTION_BLOCK

PROGRAM program0
  VAR
	IN :	BOOL;
	PT :	TIME;
	Q :	BOOL;
	func_block : TMIN;
  END_VAR
	func_block.IN  :=IN;
	func_block.PT  :=PT;
	func_block();
	Q := func_block.Q;

END_PROGRAM

CONFIGURATION Config0
	RESOURCE Res0 ON PLC
		TASK task0(INTERVAL := T#20ms,PRIORITY := 0);
		PROGRAM instance0 WITH task0 : program0;
	END_RESOURCE
END_CONFIGURATION

(* ---- 160-DWORD_TO_STRH.ST ---- *)
FUNCTION_BLOCK DWORD_TO_STRH_Block

	VAR_INPUT
		IN :	DWORD;
	END_VAR

	VAR_OUTPUT
		DWORD_TO_STRH :	STRING;
	END_VAR

	DWORD_TO_STRH:=DWORD_TO_STRING(IN);

END_FUNCTION_BLOCK

PROGRAM program0
  VAR
    LocalVar0 : DWORD;
	LocalOUT  : STRING;
	func_block : DWORD_TO_STRH_Block;
  END_VAR
	func_block.IN  := LocalVar0;
	func_block();
	LocalOUT := func_block.DWORD_TO_STRH;
END_PROGRAM

CONFIGURATION Config0
  RESOURCE Res0 ON PLC
    TASK task0(INTERVAL := T#20ms,PRIORITY := 0);
    PROGRAM instance0 WITH task0 : program0;
  END_RESOURCE
END_CONFIGURATION

(* ---- 174-R2_SET.ST ---- *)
TYPE REAL2 :

	STRUCT
		R1 : REAL;
		RX : REAL;
	END_STRUCT;

END_TYPE

FUNCTION_BLOCK R2_SET_Block

	VAR_INPUT
		X :	REAL;
	END_VAR

	VAR_OUTPUT
		R2_SET :	REAL2;
	END_VAR

	R2_SET.RX := X;
	R2_SET.R1 := 0.0;

END_FUNCTION_BLOCK

PROGRAM program0

	VAR
		X :	REAL;

        R2_SET :	REAL2;
		func_block : R2_SET_Block;
	END_VAR
	func_block.X := X;
	func_block();
	R2_SET := func_block.R2_SET;

	END_PROGRAM

CONFIGURATION Config0

	RESOURCE Res0 ON PLC
		TASK task0(INTERVAL := T#20ms,PRIORITY := 0);
		PROGRAM instance0 WITH task0 : program0;
	END_RESOURCE

END_CONFIGURATION

(* ---- 178-HEX_TO_DWORD.ST ---- *)
FUNCTION_BLOCK HEX_TO_DWORD

	VAR_INPUT
		HEX :	oscat_STRING20;
	END_VAR

	VAR_OUTPUT
		HEX_TO_DWORD :	DWORD;
	END_VAR

	VAR
		i :	INT;
		stop :	INT;
		X :	INT;
	END_VAR

	HEX_TO_DWORD := DWORD#0;
	stop := LEN(Hex);
	FOR I := 1 TO stop DO
		x := GET_CHAR(Hex,I);
		IF X > 47 AND x < 58 THEN
			HEX_TO_DWORD := SHL_DWORD(HEX_TO_DWORD,4) OR INT_TO_DWORD (X - 48);
		ELSIF X > 64 AND X < 71 THEN
			HEX_TO_DWORD := SHL_DWORD(HEX_TO_DWORD,4) OR INT_TO_DWORD (X - 55);
		ELSIF X > 96 AND X < 103 THEN
			HEX_TO_DWORD := SHL_DWORD(HEX_TO_DWORD,4) OR INT_TO_DWORD (X - 87);
		END_IF;
	END_FOR;

END_FUNCTION_BLOCK

(* ---- 18-PIN_CODE.ST ---- *)
FUNCTION_BLOCK PIN_CODE_Block

	VAR_INPUT
		CB :	BYTE;
		E :	BOOL;
		PIN :	STRING;
	END_VAR

	VAR_OUTPUT
		_TP :	BOOL;
	END_VAR

	VAR
		POS :	INT := 1;
	END_VAR

	_tp := FALSE;
	IF e THEN

		IF CB = INT_TO_BYTE(GET_CHAR(PIN,POS)) THEN
			pos := pos + 1;
			IF pos > LEN(PIN) THEN
				_TP := TRUE;
				pos := 1;
			END_IF;
		ELSE
			pos := 1;
		END_IF;
	END_IF;

END_FUNCTION_BLOCK

(* ---- 180-DEC_2.ST ---- *)
FUNCTION_BLOCK DEC_2
	VAR_INPUT
		D :	BOOL;
		A :	BOOL;
	END_VAR
	VAR_OUTPUT
		Q0 :	BOOL;
		Q1 :	BOOL;
	END_VAR
	Q0 := D AND NOT A;
	Q1 := D AND A;
END_FUNCTION_BLOCK

PROGRAM program0
  VAR
    LocalVar0 : BOOL;
	LocalVar1 : BOOL;
	LocalOUT  : BOOL;
	LocalOUT1  : BOOL;
	func_block : DEC_2;
  END_VAR
	func_block.D  := LocalVar0;
	func_block.A  := LocalVar1;
	func_block();
	LocalOUT := func_block.Q0;
	LocalOUT1 := func_block.Q1;
END_PROGRAM

CONFIGURATION Config0
  RESOURCE Res0 ON PLC
    TASK task0(INTERVAL := T#20ms,PRIORITY := 0);
    PROGRAM instance0 WITH task0 : program0;
  END_RESOURCE
END_CONFIGURATION

(* ---- 181-TOGGLE.ST ---- *)
FUNCTION_BLOCK TOGGLE

	VAR_INPUT
		CLK :	BOOL;
		RST :	BOOL;
	END_VAR

	VAR_OUTPUT
		Q :	BOOL;
	END_VAR

	VAR
		edge :	BOOL;
	END_VAR

	IF rst THEN
		Q := FALSE;
	ELSIF clk AND NOT edge THEN
		Q := NOT Q;
	END_IF;
	edge := clk;

END_FUNCTION_BLOCK

PROGRAM program0
  VAR
	CLK :	BOOL;
	RST :	BOOL;
	Q :	BOOL;
	func_block : TOGGLE;
  END_VAR
	func_block.CLK  :=CLK;
	func_block.RST  :=RST;
	func_block();
	Q := func_block.Q;

END_PROGRAM

CONFIGURATION Config0
	RESOURCE Res0 ON PLC
		TASK task0(INTERVAL := T#20ms,PRIORITY := 0);
		PROGRAM instance0 WITH task0 : program0;
	END_RESOURCE
END_CONFIGURATION

(* ---- 182-DEAD_ZONE2.ST ---- *)
FUNCTION_BLOCK DEAD_ZONE2
	VAR_INPUT
		X :	REAL;
		L :	REAL;
	END_VAR

	VAR_OUTPUT
		Y :	REAL;
	END_VAR

	IF ABS(x) > L THEN
		Y := X;
	ELSIF Y > 0.0 THEN
		Y := L;
	ELSE
		Y := -L;
	END_IF;
END_FUNCTION_BLOCK

PROGRAM program0
  VAR
    LocalVar0 : REAL;
	LocalVar1 : REAL;
	LocalOUT  : REAL;
	func_block : DEAD_ZONE2;
  END_VAR
	func_block.X  := LocalVar0;
	func_block.L  := LocalVar1;
	func_block();
	LocalOUT := func_block.Y;
END_PROGRAM

CONFIGURATION Config0
  RESOURCE Res0 ON PLC
    TASK task0(INTERVAL := T#20ms,PRIORITY := 0);
    PROGRAM instance0 WITH task0 : program0;
  END_RESOURCE
END_CONFIGURATION

(* ---- 183-V3_ABS.ST ---- *)
TYPE oscat_vector_3:
	STRUCT
		X : REAL;
		Y : REAL;
		Z : REAL;
	END_STRUCT;
END_TYPE

FUNCTION_BLOCK V3_ABS_Block

	VAR_INPUT
		A :	oscat_vector_3;
	END_VAR

	VAR_OUTPUT
		V3_ABS :	REAL;
	END_VAR

	V3_ABS := SQRT(A.X * A.X + A.Y * A.Y + A.Z * A.Z);

END_FUNCTION_BLOCK

PROGRAM program0
  	VAR
		A :	oscat_vector_3;
		V3_ABS :	REAL;
		func_block : V3_ABS_Block;
  	END_VAR
	func_block.A := A;
	func_block();
	V3_ABS := func_block.V3_ABS;
END_PROGRAM

CONFIGURATION Config0
	RESOURCE Res0 ON PLC
		TASK task0(INTERVAL := T#20ms,PRIORITY := 0);
		PROGRAM instance0 WITH task0 : program0;
	END_RESOURCE
END_CONFIGURATION

(* ---- 184-D_TRIG.ST ---- *)
FUNCTION_BLOCK D_TRIG
	VAR_INPUT
		IN :	DWORD;
	END_VAR

	VAR_OUTPUT
		Q :	BOOL;
		X :	DWORD;
	END_VAR

	VAR
		last_in :	DWORD;
	END_VAR

	Q := in <> last_in;
	X := UDINT_TO_DWORD(DWORD_TO_UDINT(in) - DWORD_TO_UDINT(last_in));
	last_in := in;
END_FUNCTION_BLOCK

PROGRAM program0
  VAR
	IN :	DWORD;

	Q :	BOOL;
	X :	DWORD;

	func_block : D_TRIG;
  END_VAR
	func_block.IN  := IN;
	func_block();
	Q := func_block.Q;
	X := func_block.X;
END_PROGRAM

CONFIGURATION Config0
  RESOURCE Res0 ON PLC
    TASK task0(INTERVAL := T#20ms,PRIORITY := 0);
    PROGRAM instance0 WITH task0 : program0;
  END_RESOURCE
END_CONFIGURATION

(* ---- 187-V3_NUL.ST ---- *)
TYPE oscat_vector_3:
	STRUCT
		X : REAL;
		Y : REAL;
		Z : REAL;
	END_STRUCT;
END_TYPE

FUNCTION_BLOCK V3_NUL_Block

	VAR_INPUT
		A :	oscat_vector_3;
	END_VAR

	VAR_OUTPUT
		V3_NUL :	BOOL;
	END_VAR

	V3_NUL := A.X = 0.0 AND A.Y = 0.0 AND A.Z = 0.0;

END_FUNCTION_BLOCK

PROGRAM program0
  	VAR
		A :	oscat_vector_3;
		V3_NUL :	BOOL;
		func_block : V3_NUL_Block;
  	END_VAR
	func_block.A := A;
	func_block();
	V3_NUL := func_block.V3_NUL;
END_PROGRAM

CONFIGURATION Config0
  RESOURCE Res0 ON PLC
    TASK task0(INTERVAL := T#20ms,PRIORITY := 0);
    PROGRAM instance0 WITH task0 : program0;
  END_RESOURCE
END_CONFIGURATION

(* ---- 189-CCON.ST ---- *)
TYPE oscat_complex :
  STRUCT
	re : REAL;
	im : REAL;
  END_STRUCT;
END_TYPE

FUNCTION_BLOCK CCON_Block

	VAR_INPUT
		X :	oscat_complex;
	END_VAR

	VAR_OUTPUT
		CCON :	oscat_complex;
	END_VAR

	CCON.re := x.re;
	CCON.im := -x.im;

END_FUNCTION_BLOCK

PROGRAM program0
  VAR
    LocalVar0 : oscat_complex;
	LocalOUT  : oscat_complex;
	func_block : CCON_Block;
  END_VAR
	func_block.X  := LocalVar0;
	func_block();
	LocalOUT := func_block.CCON;
END_PROGRAM

CONFIGURATION Config0
  RESOURCE Res0 ON PLC
    TASK task0(INTERVAL := T#20ms,PRIORITY := 0);
    PROGRAM instance0 WITH task0 : program0;
  END_RESOURCE
END_CONFIGURATION

(* ---- 190-TRIM.ST ---- *)
FUNCTION_BLOCK TRIM

	VAR_INPUT
		STR :	STRING;
	END_VAR

	VAR_OUTPUT
		TRIM3 :	STRING;
	END_VAR

	VAR
		pos :	INT;
	END_VAR

	trim3 := str;
	REPEAT
		pos := FIND(trim3,' ');
		IF pos > 0 THEN trim3 := REPLACE(trim3,'',1,pos); END_IF;
	UNTIL pos = 0 END_REPEAT;

END_FUNCTION_BLOCK

PROGRAM program0
  VAR
	STR :	STRING;

	TRIM3 :	STRING;
	func_block : TRIM;
  END_VAR
	func_block.STR  :=STR ;
	func_block();
	TRIM3 := func_block.TRIM3;

END_PROGRAM

CONFIGURATION Config0
	RESOURCE Res0 ON PLC
		TASK task0(INTERVAL := T#20ms,PRIORITY := 0);
		PROGRAM instance0 WITH task0 : program0;
	END_RESOURCE
END_CONFIGURATION

(* ---- 191-BOOL_TO_STRING.ST ---- *)
TYPE
  oscat_STRING1               : STRING(1);
END_TYPE

FUNCTION_BLOCK BOOL_TO_STRING_Block
	VAR_INPUT
		IN :	BOOL;
	END_VAR

	VAR_OUTPUT
		BOOL_TO_STRING :	oscat_STRING1;
	END_VAR

	BOOL_TO_STRING := SEL_STRING(IN,'0','1');
END_FUNCTION_BLOCK

PROGRAM program0
  VAR
    LocalVar0 : BOOL;
	LocalOUT  : oscat_STRING1;
	func_block : BOOL_TO_STRING_Block;
  END_VAR
	func_block.IN := LocalVar0;
	func_block();
	LocalOUT := func_block.BOOL_TO_STRING;

END_PROGRAM

CONFIGURATION Config0
  RESOURCE Res0 ON PLC
    TASK task0(INTERVAL := T#20ms,PRIORITY := 0);
    PROGRAM instance0 WITH task0 : program0;
  END_RESOURCE
END_CONFIGURATION

(* ---- 199-R2_MUL.ST ---- *)
TYPE REAL2 :

	STRUCT
		R1 : REAL;
		RX : REAL;
	END_STRUCT;

END_TYPE

FUNCTION_BLOCK R2_MUL_Block

	VAR_INPUT
		X :	REAL2;
		Y :	REAL;
	END_VAR

	VAR_OUTPUT
		R2_MUL :	REAL2;
	END_VAR

	R2_MUL.RX := X.RX * Y;
	R2_MUL.R1 := X.R1 * Y;

END_FUNCTION_BLOCK

PROGRAM program0

	VAR
		X :	REAL2;
		Y :	REAL;

        R2_MUL :	REAL2;
		func_block : R2_MUL_Block;
	END_VAR
	func_block.X := X;
	func_block.Y := Y;
	func_block();
	R2_MUL := func_block.R2_MUL;

	END_PROGRAM

CONFIGURATION Config0

	RESOURCE Res0 ON PLC
		TASK task0(INTERVAL := T#20ms,PRIORITY := 0);
		PROGRAM instance0 WITH task0 : program0;
	END_RESOURCE

END_CONFIGURATION

(* ---- 2-CODE.ST ---- *)
FUNCTION_BLOCK CODE_Block
	VAR_INPUT
		STR :	STRING;
		POS :	INT;
	END_VAR

	VAR_OUTPUT
		CODE :	BYTE;
	END_VAR

	IF pos < 1 OR pos > LEN(str) THEN
		CODE := BYTE#0;
		RETURN;
	ELSE
		CODE := INT_TO_BYTE(GET_CHAR(STR,POS));
	END_IF;
END_FUNCTION_BLOCK

(* ---- 201-R2_DIV.ST ---- *)
TYPE REAL2 :

	STRUCT
		R1 : REAL;
		RX : REAL;
	END_STRUCT;

END_TYPE

FUNCTION_BLOCK R2_DIV_Block

	VAR_INPUT
		X :	REAL2;
		Y :	REAL;
	END_VAR

	VAR_OUTPUT
		R2_DIV :	REAL2;
	END_VAR

	R2_DIV.RX := X.RX / Y;
	R2_DIV.R1 := X.R1 / Y;

END_FUNCTION_BLOCK

PROGRAM program0

	VAR
		X :	REAL2;
		Y :	REAL;

        R2_DIV :	REAL2;
		func_block : R2_DIV_Block;
	END_VAR
	func_block.X := X;
	func_block.Y := Y;
	func_block();
	R2_DIV := func_block.R2_DIV;

END_PROGRAM

CONFIGURATION Config0

	RESOURCE Res0 ON PLC
		TASK task0(INTERVAL := T#20ms,PRIORITY := 0);
		PROGRAM instance0 WITH task0 : program0;
	END_RESOURCE

END_CONFIGURATION

(* ---- 202-V3_REV.ST ---- *)
TYPE oscat_vector_3:
	STRUCT
		X : REAL;
		Y : REAL;
		Z : REAL;
	END_STRUCT;
END_TYPE

FUNCTION_BLOCK V3_REV_Block
	VAR_INPUT
		A :	oscat_vector_3;
	END_VAR

	VAR_OUTPUT
		V3_REV :	oscat_vector_3;
	END_VAR

	V3_REV.X := -A.X;
	V3_REV.Y := -A.Y;
	V3_REV.Z := -A.Z;

END_FUNCTION_BLOCK

PROGRAM program0
  	VAR
		A :	oscat_vector_3;
		V3_REV : oscat_vector_3;
		func_block : V3_REV_Block;
  	END_VAR
	func_block.A := A;
	func_block();
	V3_REV := func_block.V3_REV;
END_PROGRAM

CONFIGURATION Config0
  RESOURCE Res0 ON PLC
    TASK task0(INTERVAL := T#20ms,PRIORITY := 0);
    PROGRAM instance0 WITH task0 : program0;
  END_RESOURCE
END_CONFIGURATION

(* ---- 207-CODE_250.ST ---- *)
FUNCTION_BLOCK CODE_250
	VAR_INPUT
		STR :	STRING;
		POS :	INT;
	END_VAR

	VAR_OUTPUT
		CODE :	BYTE;
	END_VAR

	IF pos < 1 OR pos > LEN(str) THEN
		CODE := BYTE#0;
		RETURN;
	ELSE
		CODE := INT_TO_BYTE(GET_CHAR(STR,POS));
	END_IF;
END_FUNCTION_BLOCK

PROGRAM program0
  VAR
    LocalVar0 : STRING;
	LocalVar1 : INT;
	LocalOUT  : BYTE;
	func_block : CODE_250;
  END_VAR
	func_block.STR  := LocalVar0;
	func_block.POS  := LocalVar1;
	func_block();
	LocalOUT := func_block.CODE;
END_PROGRAM

CONFIGURATION Config0
  RESOURCE Res0 ON PLC
    TASK task0(INTERVAL := T#20ms,PRIORITY := 0);
    PROGRAM instance0 WITH task0 : program0;
  END_RESOURCE
END_CONFIGURATION

(* ---- 211-R2_ADD2.ST ---- *)
TYPE REAL2 :

	STRUCT
		R1 : REAL;
		RX : REAL;
	END_STRUCT;

END_TYPE

FUNCTION_BLOCK R2_ADD2_Block

	VAR_INPUT
		X :	REAL2;
		Y :	REAL2;
	END_VAR

	VAR_OUTPUT
		R2_ADD2 :	REAL2;
	END_VAR

	R2_ADD2.R1 := X.R1 + Y.R1;
	R2_ADD2.RX := X.RX + Y.RX;

END_FUNCTION_BLOCK

PROGRAM program0

	VAR
		X :	REAL2;
		Y :	REAL2;

        R2_ADD2 :	REAL2;
		func_block : R2_ADD2_Block;
	END_VAR
	func_block.X := X;
	func_block.Y := Y;
	func_block();
	R2_ADD2 := func_block.R2_ADD2;

END_PROGRAM

CONFIGURATION Config0

	RESOURCE Res0 ON PLC
		TASK task0(INTERVAL := T#20ms,PRIORITY := 0);
		PROGRAM instance0 WITH task0 : program0;
	END_RESOURCE

END_CONFIGURATION

(* ---- 214-MIRROR.ST ---- *)
FUNCTION_BLOCK MIRROR_Block

	VAR_INPUT
		STR :	STRING;
	END_VAR

	VAR_OUTPUT
		MIRROR :	STRING;
	END_VAR

	VAR
		i :	INT;
		st_temp :	STRING;
	END_VAR

	mirror := '';
	i := LEN(str);
	WHILE i > 0 DO
	st_temp := MID(str,1,i);
	mirror := CONCAT(mirror,st_temp);
	i := i -1;
	END_WHILE;

END_FUNCTION_BLOCK

PROGRAM program0

	VAR
		STR :	STRING;
		MIRROR :	STRING;
		func_block : MIRROR_Block;
	END_VAR
	func_block.STR := STR;
	func_block();
	MIRROR  := func_block.MIRROR;

END_PROGRAM

CONFIGURATION Config0

	RESOURCE Res0 ON PLC
		TASK task0(INTERVAL := T#20ms,PRIORITY := 0);
		PROGRAM instance0 WITH task0 : program0;
	END_RESOURCE

END_CONFIGURATION

(* ---- 215-CSET.ST ---- *)
TYPE oscat_complex :
  STRUCT
	re : REAL;
	im : REAL;
  END_STRUCT;
END_TYPE

FUNCTION_BLOCK CSET_Block
	VAR_INPUT
		RE :	REAL;
		IM :	REAL;
	END_VAR

	VAR_OUTPUT
		CSET :	oscat_complex;
	END_VAR

	CSET.re := RE;
	CSET.im := IM;
END_FUNCTION_BLOCK

PROGRAM program0
  VAR
    LocalVar0 : REAL;
	LocalVar1 : REAL;
	LocalOUT  : oscat_complex;
	func_block : CSET_Block;
  END_VAR
	func_block.RE  := LocalVar0;
	func_block.IM  := LocalVar1;
	func_block();
	LocalOUT := func_block.CSET;
END_PROGRAM

CONFIGURATION Config0
  RESOURCE Res0 ON PLC
    TASK task0(INTERVAL := T#20ms,PRIORITY := 0);
    PROGRAM instance0 WITH task0 : program0;
  END_RESOURCE
END_CONFIGURATION

(* ---- 217-CPOL.ST ---- *)
TYPE oscat_complex :
  STRUCT
	re : REAL;
	im : REAL;
  END_STRUCT;
END_TYPE

FUNCTION_BLOCK CPOL_Block
	VAR_INPUT
		L :	REAL;
		A :	REAL;
	END_VAR

	VAR_OUTPUT
		CPOL :	oscat_complex;
	END_VAR

	CPOL.re := L * COS(A);
	CPOL.im := L * SIN(A);
END_FUNCTION_BLOCK

PROGRAM program0
  VAR
    LocalVar0 : REAL;
	LocalVar1 : REAL;
	CPOL  : oscat_complex;
	func_block : CPOL_Block;
  END_VAR
	func_block.L  := LocalVar0;
	func_block.A  := LocalVar1;
	func_block();
	CPOL := func_block.CPOL;
END_PROGRAM

CONFIGURATION Config0
  RESOURCE Res0 ON PLC
    TASK task0(INTERVAL := T#20ms,PRIORITY := 0);
    PROGRAM instance0 WITH task0 : program0;
  END_RESOURCE
END_CONFIGURATION

(* ---- 219-LTCH.ST ---- *)
FUNCTION_BLOCK LTCH_Block

	VAR_INPUT
		D :	BOOL;
		L :	BOOL;
		RST :	BOOL;
	END_VAR

	VAR_OUTPUT
		Q :	BOOL;
	END_VAR

	IF rst THEN				(* if asynchronous reset then Q=0 *)
		Q := FALSE;
	ELSIF L THEN			(* latch is transparent *)
		Q := D;
	END_IF;

END_FUNCTION_BLOCK

PROGRAM program0

	VAR
		D :	BOOL;
		L :	BOOL;
		RST :	BOOL;

		Q :	BOOL;

		func_block : LTCH_Block;
	END_VAR
	func_block.D := D;
	func_block.L := L;
	func_block.RST := RST;

	func_block();
	Q := func_block.Q;

END_PROGRAM

CONFIGURATION Config0

	RESOURCE Res0 ON PLC
		TASK task0(INTERVAL := T#20ms,PRIORITY := 0);
		PROGRAM instance0 WITH task0 : program0;
	END_RESOURCE

END_CONFIGURATION

(* ---- 220-IS_NUM.ST ---- *)
FUNCTION_BLOCK IS_NUM_Block

	VAR_INPUT
		STR :	STRING;
	END_VAR

	VAR_OUTPUT
		IS_NUM :	BOOL;
	END_VAR

	VAR
		pos :	INT;
		I :	INT;
	END_VAR

	I := LEN(str);
	FOR pos := 1 TO I DO
		IF NOT ISC_NUM(INT_TO_BYTE(GET_CHAR(str,pos))) THEN
			IS_NUM := FALSE;
			RETURN;
		END_IF;
	END_FOR;
	IS_NUM := I>0;

END_FUNCTION_BLOCK

PROGRAM program0

	VAR
		STR :	STRING;
		IS_NUM :	BOOL;
		func_block : IS_NUM_Block;
	END_VAR
	func_block.STR := STR;
	func_block();
	IS_NUM := func_block.IS_NUM;

END_PROGRAM

CONFIGURATION Config0

	RESOURCE Res0 ON PLC
		TASK task0(INTERVAL := T#20ms,PRIORITY := 0);
		PROGRAM instance0 WITH task0 : program0;
	END_RESOURCE

END_CONFIGURATION

(* ---- 222-R2_ABS.ST ---- *)
TYPE REAL2 :

	STRUCT
		R1 : REAL;
		RX : REAL;
	END_STRUCT;

END_TYPE

FUNCTION_BLOCK R2_ABS_Block

	VAR_INPUT
		X :	REAL2;
	END_VAR

	VAR_OUTPUT
		R2_ABS :	REAL2;
	END_VAR

	IF X.RX >= 0.0 THEN
		R2_ABS.RX := X.RX;
		R2_ABS.R1 := X.R1;
	ELSE
		R2_ABS.RX := -X.RX;
		R2_ABS.R1 := -X.R1;
	END_IF;

END_FUNCTION_BLOCK

PROGRAM program0

	VAR
		X :	REAL2;

        R2_ABS :	REAL2;
		func_block : R2_ABS_Block;
	END_VAR
	func_block.X := X;
	func_block();
	R2_ABS := func_block.R2_ABS;

END_PROGRAM

CONFIGURATION Config0

	RESOURCE Res0 ON PLC
		TASK task0(INTERVAL := T#20ms,PRIORITY := 0);
		PROGRAM instance0 WITH task0 : program0;
	END_RESOURCE

END_CONFIGURATION

(* ---- 223-DEBOUNCE.ST ---- *)
FUNCTION_BLOCK DEBOUNCE_Block

	VAR_INPUT
		IN :	BOOL;
		TD :	TIME;
		PM :	BOOL;
	END_VAR

	VAR_OUTPUT
		Q :	BOOL;
	END_VAR

	VAR
		deb :	TOF;
	END_VAR

	IF NOT deb.Q AND IN THEN
		Q := TRUE;
	ELSIF NOT PM THEN
		Q := deb.Q;
	ELSE
		Q := FALSE;
	END_IF;

END_FUNCTION_BLOCK

PROGRAM program0
	VAR
		IN :	BOOL;
		TD :	TIME;
		PM :	BOOL;
		Q :	BOOL;

		func_block : DEBOUNCE_Block;
	END_VAR
	func_block.IN := IN;
	func_block.TD := TD;
	func_block.PM := PM ;

	func_block();
	Q  := func_block.Q;
END_PROGRAM

CONFIGURATION Config0
	RESOURCE Res0 ON PLC
		TASK task0(INTERVAL := T#20ms,PRIORITY := 0);
		PROGRAM instance0 WITH task0 : program0;
	END_RESOURCE
END_CONFIGURATION

(* ---- 227-V3_DPRO.ST ---- *)
TYPE oscat_vector_3:
	STRUCT
		X : REAL;
		Y : REAL;
		Z : REAL;
	END_STRUCT;
END_TYPE

FUNCTION_BLOCK V3_DPRO_Block

	VAR_INPUT
		A :	oscat_vector_3;
		B :	oscat_vector_3;
	END_VAR

	VAR_OUTPUT
		V3_DPRO :	REAL;
	END_VAR

	V3_DPRO := A.X * B.X + A.Y * B.Y + A.Z * B.Z;

END_FUNCTION_BLOCK

PROGRAM program0
  	VAR
		A :	oscat_vector_3;
		B :	oscat_vector_3;
		V3_DPRO : REAL;
		func_block : V3_DPRO_Block;
  	END_VAR
	func_block.A := A;
	func_block.B := B;
	func_block();
	V3_DPRO := func_block.V3_DPRO;
END_PROGRAM

CONFIGURATION Config0
  RESOURCE Res0 ON PLC
    TASK task0(INTERVAL := T#20ms,PRIORITY := 0);
    PROGRAM instance0 WITH task0 : program0;
  END_RESOURCE
END_CONFIGURATION

(* ---- 228-SH.ST ---- *)
FUNCTION_BLOCK SH_Block

	VAR_INPUT
		IN :	REAL;
		CLK :	BOOL;
	END_VAR

	VAR_OUTPUT
		OUT :	REAL;
		TRIG :	BOOL;
	END_VAR

	VAR
		edge :	BOOL;
	END_VAR

	IF clk AND NOT edge THEN
		out := in;
		trig := TRUE;
	ELSE
		trig := FALSE;
	END_IF;
	edge := clk;

END_FUNCTION_BLOCK

PROGRAM program0

	VAR
		IN :	REAL;
		CLK :	BOOL;
		OUT :	REAL;
		TRIG :	BOOL;
		func_block : SH_Block;
	END_VAR
		func_block.IN  :=IN;
		func_block.CLK  :=CLK;
		func_block();
		OUT := func_block.OUT;
		TRIG := func_block.TRIG;

END_PROGRAM

CONFIGURATION Config0
	RESOURCE Res0 ON PLC
		TASK task0(INTERVAL := T#20ms,PRIORITY := 0);
		PROGRAM instance0 WITH task0 : program0;
	END_RESOURCE
END_CONFIGURATION

(* ---- 232-TREND.ST ---- *)
FUNCTION_BLOCK TREND

	VAR_INPUT
		X :	REAL;
	END_VAR

	VAR_OUTPUT
		Q :	BOOL;
		TU :	BOOL;
		TD :	BOOL;
		D :	REAL;
	END_VAR

	VAR
		last_x :	REAL;
	END_VAR

	TU := X > last_X;
	TD := X < last_X;
	Q := TU OR TD;
	D := X - LAST_X;

	last_X := X;

END_FUNCTION_BLOCK

PROGRAM program0
  VAR
	X :	REAL;
	Q :	BOOL;
	TU :	BOOL;
	TD :	BOOL;
	D :	REAL;
	func_block : TREND;
  END_VAR
	func_block.X  :=X ;
	func_block();
	Q := func_block.Q;
	TU := func_block.TU;
	TD := func_block.TD;
	D := func_block.D;
END_PROGRAM

CONFIGURATION Config0
	RESOURCE Res0 ON PLC
		TASK task0(INTERVAL := T#20ms,PRIORITY := 0);
		PROGRAM instance0 WITH task0 : program0;
	END_RESOURCE
END_CONFIGURATION

(* ---- 233-CEXP.ST ---- *)
TYPE oscat_complex :
  STRUCT
	re : REAL;
	im : REAL;
  END_STRUCT;
END_TYPE

FUNCTION_BLOCK CEXP_Block
	VAR_INPUT
		X :	oscat_complex;
	END_VAR

	VAR_OUTPUT
		CEXP :	oscat_complex;
	END_VAR

	VAR
		Temp :	REAL;
	END_VAR

	temp := EXP(X.re);
	CEXP.re := temp * COS(X.im);
	CEXP.im := temp * SIN(X.im);

END_FUNCTION_BLOCK

PROGRAM program0
  VAR
    LocalVar0 : oscat_complex;
	LocalOUT  : oscat_complex;
	func_block : CEXP_Block;
  END_VAR
	func_block.X  := LocalVar0;
	func_block();
	LocalOUT := func_block.CEXP;
END_PROGRAM

CONFIGURATION Config0
  RESOURCE Res0 ON PLC
    TASK task0(INTERVAL := T#20ms,PRIORITY := 0);
    PROGRAM instance0 WITH task0 : program0;
  END_RESOURCE
END_CONFIGURATION

(* ---- 235-V3_SMUL.ST ---- *)
TYPE oscat_vector_3:
	STRUCT
		X : REAL;
		Y : REAL;
		Z : REAL;
	END_STRUCT;
END_TYPE

FUNCTION_BLOCK V3_SMUL_Block
	VAR_INPUT
		A :	oscat_vector_3;
		M :	REAL;
	END_VAR

	VAR_OUTPUT
		V3_SMUL :	oscat_vector_3;
	END_VAR

	V3_SMUL.X := A.X * M;
	V3_SMUL.Y := A.Y * M;
	V3_SMUL.Z := A.Z * M;
END_FUNCTION_BLOCK

PROGRAM program0
  	VAR
		A :	oscat_vector_3;
		M :	REAL;
		V3_SMUL :	oscat_vector_3;
		func_block : V3_SMUL_Block;
  	END_VAR
	func_block.A := A;
	func_block.M := M;
	func_block();
	V3_SMUL := func_block.V3_SMUL;
END_PROGRAM

CONFIGURATION Config0
	RESOURCE Res0 ON PLC
		TASK task0(INTERVAL := T#20ms,PRIORITY := 0);
		PROGRAM instance0 WITH task0 : program0;
	END_RESOURCE
END_CONFIGURATION

(* ---- 236-F_POLY.ST ---- *)
TYPE
  oscat_arr_0_7               : ARRAY [0..7]    OF REAL;
END_TYPE

FUNCTION_BLOCK F_POLY_Block
	VAR_INPUT
		X :	REAL;
		C :	oscat_arr_0_7;
	END_VAR

	VAR_OUTPUT
		F_POLY :	REAL;
	END_VAR

	F_POLY := ((((((( c[7] * x + c[6] ) * x + c[5] ) * x + c[4] ) * x + c[3] ) * x + c[2] ) * x + c[1] ) * x + c[0] ) ;

END_FUNCTION_BLOCK

PROGRAM program0
	VAR
		X :	REAL;
		C :	oscat_arr_0_7;

		F_POLY :	REAL;

		func_block : F_POLY_Block;
	END_VAR
	func_block.X := X;
	func_block.C := C;
	func_block();
	F_POLY  := func_block.F_POLY;
END_PROGRAM

CONFIGURATION Config0
	RESOURCE Res0 ON PLC
		TASK task0(INTERVAL := T#20ms,PRIORITY := 0);
		PROGRAM instance0 WITH task0 : program0;
	END_RESOURCE
END_CONFIGURATION

(* ---- 238-CABS.ST ---- *)
TYPE oscat_complex :
  STRUCT
	re : REAL;
	im : REAL;
  END_STRUCT;
END_TYPE

FUNCTION HYPOT:REAL
	VAR_INPUT
		X :	REAL;
		Y :	REAL;
	END_VAR

	HYPOT := SQRT(x*x + y*y);
END_FUNCTION

FUNCTION_BLOCK CABS_Block
	VAR_INPUT
		X :	oscat_complex;
	END_VAR

	VAR_OUTPUT
		CABS :	REAL;
	END_VAR

	CABS := HYPOT(x.re, x.im);

END_FUNCTION_BLOCK

PROGRAM program0
  VAR
    LocalVar0 : oscat_complex;
	LocalOUT  : REAL;
	func_block : CABS_Block;
  END_VAR
	func_block.X  := LocalVar0;
	func_block();
	LocalOUT := func_block.CABS;

END_PROGRAM

CONFIGURATION Config0
  RESOURCE Res0 ON PLC
    TASK task0(INTERVAL := T#20ms,PRIORITY := 0);
    PROGRAM instance0 WITH task0 : program0;
  END_RESOURCE
END_CONFIGURATION

(* ---- 240-CSUB.ST ---- *)
TYPE oscat_complex :
  STRUCT
	re : REAL;
	im : REAL;
  END_STRUCT;
END_TYPE

FUNCTION_BLOCK CSUB_Block
	VAR_INPUT
		X :	oscat_complex;
		Y :	oscat_complex;
	END_VAR

	VAR_OUTPUT
		CSUB :	oscat_complex;
	END_VAR

	CSUB.re := X.re - Y.re;
	CSUB.im := X.im - Y.im;
END_FUNCTION_BLOCK

PROGRAM program0
  VAR
    LocalVar0 : oscat_complex;
	LocalVar1 : oscat_complex;
	LocalOUT  : oscat_complex;
	func_block : CSUB_Block;
  END_VAR
	func_block.X  := LocalVar0;
	func_block.Y  := LocalVar0;
	func_block();
	LocalOUT := func_block.CSUB;
END_PROGRAM

CONFIGURATION Config0
  RESOURCE Res0 ON PLC
    TASK task0(INTERVAL := T#20ms,PRIORITY := 0);
    PROGRAM instance0 WITH task0 : program0;
  END_RESOURCE
END_CONFIGURATION

(* ---- 241-FF_DRE.ST ---- *)
FUNCTION_BLOCK FF_DRE
	VAR_INPUT
		SET :	BOOL;
		D :	BOOL;
		CLK :	BOOL;
		RST :	BOOL;
	END_VAR

	VAR_OUTPUT
		Q :	BOOL;
	END_VAR

	VAR
		edge :	BOOL;
	END_VAR

	IF rst OR set THEN
		Q := NOT rst;
	ELSIF clk AND NOT edge THEN
		Q := D;
	END_IF;
	edge := CLK;

END_FUNCTION_BLOCK

PROGRAM program0
  VAR
	SET :	BOOL;
	D   :	BOOL;
	CLK :	BOOL;
	RST :	BOOL;

	Q :	BOOL;

	func_block : FF_DRE;
  END_VAR
	func_block.SET:=SET;
	func_block.D  :=D  ;
	func_block.CLK:=CLK;
	func_block.RST:=RST;
	func_block();
	Q:= func_block.Q;
END_PROGRAM

CONFIGURATION Config0
  RESOURCE Res0 ON PLC
    TASK task0(INTERVAL := T#20ms,PRIORITY := 0);
    PROGRAM instance0 WITH task0 : program0;
  END_RESOURCE
END_CONFIGURATION

(* ---- 243-DELAY_4.ST ---- *)
FUNCTION_BLOCK DELAY_4

	VAR_INPUT
		IN :	REAL;
	END_VAR

	VAR_OUTPUT
		OUT1 :	REAL;
		OUT2 :	REAL;
		OUT3 :	REAL;
		OUT4 :	REAL;
	END_VAR

	VAR
		temp :	REAL;
	END_VAR

	out4 := out3;
	out3 := out2;
	out2 := out1;
	out1 := temp;
	temp := in;

END_FUNCTION_BLOCK

PROGRAM program0
  VAR
	IN :	REAL;

	OUT1 :	REAL;
	OUT2 :	REAL;
	OUT3 :	REAL;
	OUT4 :	REAL;
	func_block : DELAY_4;
  END_VAR
	func_block.IN  := IN;
	func_block();
	OUT1:= func_block.OUT1;
	OUT2:= func_block.OUT2;
	OUT3:= func_block.OUT3;
	OUT4:= func_block.OUT4;
END_PROGRAM

CONFIGURATION Config0
  RESOURCE Res0 ON PLC
    TASK task0(INTERVAL := T#20ms,PRIORITY := 0);
    PROGRAM instance0 WITH task0 : program0;
  END_RESOURCE
END_CONFIGURATION

(* ---- 244-TRIME.ST ---- *)
FUNCTION_BLOCK TRIME_Block
	VAR_INPUT
		STR :	STRING;
	END_VAR

	VAR_OUTPUT
		TRIME :	STRING;
	END_VAR

	TRIME := str;
	IF LEN(TRIME) < 1 THEN RETURN; END_IF;

	WHILE (GET_CHAR(TRIME,1) = 32) DO
		TRIME := DELETE(TRIME,1,1);
	END_WHILE;

	WHILE (GET_CHAR(TRIME,LEN(TRIME)) = 32) DO
		TRIME := DELETE(TRIME,1,LEN(TRIME));
	END_WHILE;

END_FUNCTION_BLOCK

PROGRAM program0
  	VAR
		INPUT_STR :	STRING;
		OUTPUT_TRIME : STRING;
		func_block : TRIME_Block;
  	END_VAR
	func_block.STR := INPUT_STR;
	func_block();
	OUTPUT_TRIME := func_block.TRIME;
END_PROGRAM

CONFIGURATION Config0
	RESOURCE Res0 ON PLC
		TASK task0(INTERVAL := T#20ms,PRIORITY := 0);
		PROGRAM instance0 WITH task0 : program0;
	END_RESOURCE
END_CONFIGURATION

(* ---- 245-CADD.ST ---- *)
TYPE oscat_complex :
  STRUCT
	re : REAL;
	im : REAL;
  END_STRUCT;
END_TYPE

FUNCTION_BLOCK CADD_Block

	VAR_INPUT
		X :	oscat_complex;
		Y :	oscat_complex;
	END_VAR

	VAR_OUTPUT
		CADD :	oscat_complex;
	END_VAR

	CADD.re := x.re + y.re;
	CADD.im := x.im + y.im;

END_FUNCTION_BLOCK

PROGRAM program0
  VAR
    LocalVar0 : oscat_complex;
	LocalVar1 : oscat_complex;
	LocalOUT  : oscat_complex;
	func_block : CADD_Block;
  END_VAR
	func_block.X  := LocalVar0;
	func_block.Y  := LocalVar0;
	func_block();
	LocalOUT := func_block.CADD;
END_PROGRAM

CONFIGURATION Config0
  RESOURCE Res0 ON PLC
    TASK task0(INTERVAL := T#20ms,PRIORITY := 0);
    PROGRAM instance0 WITH task0 : program0;
  END_RESOURCE
END_CONFIGURATION

(* ---- 247-R2_ADD.ST ---- *)
TYPE REAL2 :

	STRUCT
		R1 : REAL;
		RX : REAL;
	END_STRUCT;

END_TYPE

FUNCTION_BLOCK R2_ADD_Block

	VAR_INPUT
		X :	REAL2;
		Y :	REAL;
	END_VAR

	VAR_OUTPUT
		R2_ADD :	REAL2;
	END_VAR

	VAR
		temp :	REAL;
	END_VAR

	temp := X.RX;
	R2_ADD.RX := Y + X.R1 + X.RX;
	R2_ADD.R1 := temp - R2_ADD.RX + Y + X.R1;

END_FUNCTION_BLOCK

PROGRAM program0

	VAR
		X :	REAL2;
		Y :	REAL;

        R2_ADD :	REAL2;
		func_block : R2_ADD_Block;
	END_VAR
	func_block.X := X;
	func_block.Y := Y;
	func_block();
	R2_ADD := func_block.R2_ADD;

END_PROGRAM

CONFIGURATION Config0

	RESOURCE Res0 ON PLC
		TASK task0(INTERVAL := T#20ms,PRIORITY := 0);
		PROGRAM instance0 WITH task0 : program0;
	END_RESOURCE

END_CONFIGURATION

(* ---- 249-V3_ADD.ST ---- *)
TYPE oscat_vector_3:
	STRUCT
		X : REAL;
		Y : REAL;
		Z : REAL;
	END_STRUCT;
END_TYPE

FUNCTION_BLOCK V3_ADD_Block
	VAR_INPUT
		A :	oscat_vector_3;
		B :	oscat_vector_3;
	END_VAR

	VAR_OUTPUT
		V3_ADD :	oscat_vector_3;
	END_VAR

	V3_ADD.X := A.X + B.X;
	V3_ADD.Y := A.Y + B.Y;
	V3_ADD.Z := A.Z + B.Z;

END_FUNCTION_BLOCK

PROGRAM program0
  	VAR
		A :	oscat_vector_3;
		B :	oscat_vector_3;
		V3_ADD :	oscat_vector_3;
		func_block : V3_ADD_Block;
  	END_VAR
	func_block.A := A;
	func_block.B := B;
	func_block();
	V3_ADD := func_block.V3_ADD;
END_PROGRAM

CONFIGURATION Config0
  RESOURCE Res0 ON PLC
    TASK task0(INTERVAL := T#20ms,PRIORITY := 0);
    PROGRAM instance0 WITH task0 : program0;
  END_RESOURCE
END_CONFIGURATION
